    CONST robtarget Target_Nom_Rint_40:=[[-62.519469,-32.68026,0],[0.707106781,0,0,0.707106781],[0,0,0,0],[9E+09,9E+09,9E+09,9E+09,9E+09,9E+09]];
    CONST robtarget Target_Nom_Rint_50:=[[-62.519469,-22.091371,0],[0.707106781,0,0,0.707106781],[0,0,0,0],[9E+09,9E+09,9E+09,9E+09,9E+09,9E+09]];
    CONST robtarget Target_Nom_Rint_60:=[[-87.445335,-22.18424,0],[0.707106781,0,0,0.707106781],[0,0,0,0],[9E+09,9E+09,9E+09,9E+09,9E+09,9E+09]];
    CONST robtarget Target_Nom_Rint_70:=[[-87.50619,-27.43225,0],[0.707106781,0,0,0.707106781],[0,0,0,0],[9E+09,9E+09,9E+09,9E+09,9E+09,9E+09]];
    CONST robtarget Target_Nom_Rint_80:=[[-87.50619,-27.43225,-20],[0.707106781,0,0,0.707106781],[0,0,0,0],[9E+09,9E+09,9E+09,9E+09,9E+09,9E+09]];
    !***********************************************************

    !Dise?o de la parte frontal
    !***********************************************************
    !Punto para acomodar orientaci?n del defector
    CONST robtarget Target_Frente_10:=[[212.749496796,-44.184,-87.888947338],[0.627211375,-0.326505577,-0.326505577,0.627211375],[0,0,0,0],[9E+09,9E+09,9E+09,9E+09,9E+09,9E+09]];
    CONST robtarget Target_Frente_20:=[[196.247119583,-40.184,-39.636157587],[0.428395846,-0.281546356,-0.169146611,0.841782675],[0,0,0,0],[9E+09,9E+09,9E+09,9E+09,9E+09,9E+09]];
    !***********************************************************
    !Dibujo de chip
    CONST robtarget Target_DibChip_10:=[[143.048,-41.184,47.089],[0.595801453,-0.480725183,-0.403998863,0.500708343],[0,0,0,0],[9E+09,9E+09,9E+09,9E+09,9E+09,9E+09]];
    CONST robtarget Target_DibChip_20:=[[123.048,-31.184,47.089],[0.595801453,-0.480725183,-0.403998863,0.500708343],[0,0,0,0],[9E+09,9E+09,9E+09,9E+09,9E+09,9E+09]];
    CONST robtarget Target_DibChip_30:=[[122.19,-34.343,47.089],[0.595801453,-0.480725183,-0.403998863,0.500708343],[0,0,0,0],[9E+09,9E+09,9E+09,9E+09,9E+09,9E+09]];
    CONST robtarget Target_DibChip_40:=[[122.19,-34.343,43.815],[0.595801453,-0.480725183,-0.403998863,0.500708343],[0,0,0,0],[9E+09,9E+09,9E+09,9E+09,9E+09,9E+09]];
    CONST robtarget Target_DibChip_50:=[[122.19,-34.343,47.089],[0.595801453,-0.480725183,-0.403998863,0.500708343],[0,0,0,0],[9E+09,9E+09,9E+09,9E+09,9E+09,9E+09]];
    CONST robtarget Target_DibChip_60:=[[119.685,-42.135,47.089],[0.595801453,-0.480725183,-0.403998863,0.500708343],[0,0,0,0],[9E+09,9E+09,9E+09,9E+09,9E+09,9E+09]];
    CONST robtarget Target_DibChip_70:=[[119.685,-42.135,43.815],[0.595801453,-0.480725183,-0.403998863,0.500708343],[0,0,0,0],[9E+09,9E+09,9E+09,9E+09,9E+09,9E+09]];
    CONST robtarget Target_DibChip_80:=[[119.685,-42.135,47.089],[0.595801453,-0.480725183,-0.403998863,0.500708343],[0,0,0,0],[9E+09,9E+09,9E+09,9E+09,9E+09,9E+09]];
    CONST robtarget Target_DibChip_90:=[[116.675,-49.746,47.089],[0.595801453,-0.480725183,-0.403998863,0.500708343],[0,0,0,0],[9E+09,9E+09,9E+09,9E+09,9E+09,9E+09]];
    CONST robtarget Target_DibChip_100:=[[116.675,-49.746,43.815],[0.595801453,-0.480725183,-0.403998863,0.500708343],[0,0,0,0],[9E+09,9E+09,9E+09,9E+09,9E+09,9E+09]];
    CONST robtarget Target_DibChip_110:=[[116.675,-49.746,47.089],[0.595801453,-0.480725183,-0.403998863,0.500708343],[0,0,0,0],[9E+09,9E+09,9E+09,9E+09,9E+09,9E+09]];
    CONST robtarget Target_DibChip_120:=[[115.333,-52.732,47.089],[0.595801453,-0.480725183,-0.403998863,0.500708343],[0,0,0,0],[9E+09,9E+09,9E+09,9E+09,9E+09,9E+09]];
    CONST robtarget Target_DibChip_130:=[[113.824,-55.86,48.528],[0.595801453,-0.480725183,-0.403998863,0.500708343],[0,0,0,0],[9E+09,9E+09,9E+09,9E+09,9E+09,9E+09]];
    CONST robtarget Target_DibChip_140:=[[113.174,-57.143,52.001],[0.595801453,-0.480725183,-0.403998863,0.500708343],[0,0,0,0],[9E+09,9E+09,9E+09,9E+09,9E+09,9E+09]];
    CONST robtarget Target_DibChip_150:=[[113.174,-57.143,55.275],[0.595801453,-0.480725183,-0.403998863,0.500708343],[0,0,0,0],[9E+09,9E+09,9E+09,9E+09,9E+09,9E+09]];
    CONST robtarget Target_DibChip_160:=[[111.639,-60.035,55.275],[0.595801453,-0.480725183,-0.403998863,0.500708343],[0,0,0,0],[9E+09,9E+09,9E+09,9E+09,9E+09,9E+09]];
    CONST robtarget Target_DibChip_170:=[[113.174,-57.143,55.275],[0.595801453,-0.480725183,-0.403998863,0.500708343],[0,0,0,0],[9E+09,9E+09,9E+09,9E+09,9E+09,9E+09]];
    CONST robtarget Target_DibChip_180:=[[113.174,-57.143,63.46],[0.595801453,-0.480725183,-0.403998863,0.500708343],[0,0,0,0],[9E+09,9E+09,9E+09,9E+09,9E+09,9E+09]];
    CONST robtarget Target_DibChip_190:=[[111.639,-60.035,63.46],[0.595801453,-0.480725183,-0.403998863,0.500708343],[0,0,0,0],[9E+09,9E+09,9E+09,9E+09,9E+09,9E+09]];
    CONST robtarget Target_DibChip_200:=[[113.174,-57.143,63.46],[0.595801453,-0.480725183,-0.403998863,0.500708343],[0,0,0,0],[9E+09,9E+09,9E+09,9E+09,9E+09,9E+09]];
    CONST robtarget Target_DibChip_210:=[[113.174,-57.143,71.646],[0.595801453,-0.480725183,-0.403998863,0.500708343],[0,0,0,0],[9E+09,9E+09,9E+09,9E+09,9E+09,9E+09]];
    CONST robtarget Target_DibChip_220:=[[111.639,-60.035,71.646],[0.595801453,-0.480725183,-0.403998863,0.500708343],[0,0,0,0],[9E+09,9E+09,9E+09,9E+09,9E+09,9E+09]];
    CONST robtarget Target_DibChip_230:=[[113.174,-57.143,71.646],[0.595801453,-0.480725183,-0.403998863,0.500708343],[0,0,0,0],[9E+09,9E+09,9E+09,9E+09,9E+09,9E+09]];
    CONST robtarget Target_DibChip_240:=[[113.174,-57.143,74.92],[0.595801453,-0.480725183,-0.403998863,0.500708343],[0,0,0,0],[9E+09,9E+09,9E+09,9E+09,9E+09,9E+09]];
    CONST robtarget Target_DibChip_250:=[[113.824,-55.86,78.393],[0.595801453,-0.480725183,-0.403998863,0.500708343],[0,0,0,0],[9E+09,9E+09,9E+09,9E+09,9E+09,9E+09]];
    CONST robtarget Target_DibChip_260:=[[115.333,-52.732,79.832],[0.595801453,-0.480725183,-0.403998863,0.500708343],[0,0,0,0],[9E+09,9E+09,9E+09,9E+09,9E+09,9E+09]];
    CONST robtarget Target_DibChip_270:=[[116.675,-49.746,79.832],[0.595801453,-0.480725183,-0.403998863,0.500708343],[0,0,0,0],[9E+09,9E+09,9E+09,9E+09,9E+09,9E+09]];
    CONST robtarget Target_DibChip_280:=[[116.675,-49.746,83.106],[0.595801453,-0.480725183,-0.403998863,0.500708343],[0,0,0,0],[9E+09,9E+09,9E+09,9E+09,9E+09,9E+09]];
    CONST robtarget Target_DibChip_290:=[[116.675,-49.746,79.832],[0.595801453,-0.480725183,-0.403998863,0.500708343],[0,0,0,0],[9E+09,9E+09,9E+09,9E+09,9E+09,9E+09]];
    CONST robtarget Target_DibChip_300:=[[119.685,-42.135,79.832],[0.595801453,-0.480725183,-0.403998863,0.500708343],[0,0,0,0],[9E+09,9E+09,9E+09,9E+09,9E+09,9E+09]];
    CONST robtarget Target_DibChip_310:=[[119.685,-42.135,83.106],[0.595801453,-0.480725183,-0.403998863,0.500708343],[0,0,0,0],[9E+09,9E+09,9E+09,9E+09,9E+09,9E+09]];
    CONST robtarget Target_DibChip_320:=[[119.685,-42.135,79.832],[0.595801453,-0.480725183,-0.403998863,0.500708343],[0,0,0,0],[9E+09,9E+09,9E+09,9E+09,9E+09,9E+09]];
    CONST robtarget Target_DibChip_330:=[[122.19,-34.343,79.832],[0.595801453,-0.480725183,-0.403998863,0.500708343],[0,0,0,0],[9E+09,9E+09,9E+09,9E+09,9E+09,9E+09]];
    CONST robtarget Target_DibChip_340:=[[122.19,-34.343,83.106],[0.595801453,-0.480725183,-0.403998863,0.500708343],[0,0,0,0],[9E+09,9E+09,9E+09,9E+09,9E+09,9E+09]];
    CONST robtarget Target_DibChip_350:=[[122.19,-34.343,79.832],[0.595801453,-0.480725183,-0.403998863,0.500708343],[0,0,0,0],[9E+09,9E+09,9E+09,9E+09,9E+09,9E+09]];
    CONST robtarget Target_DibChip_360:=[[123.048,-31.184,79.832],[0.595801453,-0.480725183,-0.403998863,0.500708343],[0,0,0,0],[9E+09,9E+09,9E+09,9E+09,9E+09,9E+09]];
    CONST robtarget Target_DibChip_370:=[[123.867,-27.809,78.393],[0.595801453,-0.480725183,-0.403998863,0.500708343],[0,0,0,0],[9E+09,9E+09,9E+09,9E+09,9E+09,9E+09]];
    CONST robtarget Target_DibChip_380:=[[124.179,-26.405,74.92],[0.595801453,-0.480725183,-0.403998863,0.500708343],[0,0,0,0],[9E+09,9E+09,9E+09,9E+09,9E+09,9E+09]];
    CONST robtarget Target_DibChip_390:=[[124.179,-26.405,71.646],[0.595801453,-0.480725183,-0.403998863,0.500708343],[0,0,0,0],[9E+09,9E+09,9E+09,9E+09,9E+09,9E+09]];
    CONST robtarget Target_DibChip_400:=[[124.829,-23.196,71.646],[0.595801453,-0.480725183,-0.403998863,0.500708343],[0,0,0,0],[9E+09,9E+09,9E+09,9E+09,9E+09,9E+09]];
    CONST robtarget Target_DibChip_410:=[[124.179,-26.405,71.646],[0.595801453,-0.480725183,-0.403998863,0.500708343],[0,0,0,0],[9E+09,9E+09,9E+09,9E+09,9E+09,9E+09]];
    CONST robtarget Target_DibChip_420:=[[124.179,-26.405,63.46],[0.595801453,-0.480725183,-0.403998863,0.500708343],[0,0,0,0],[9E+09,9E+09,9E+09,9E+09,9E+09,9E+09]];
    CONST robtarget Target_DibChip_430:=[[124.829,-23.196,63.46],[0.595801453,-0.480725183,-0.403998863,0.500708343],[0,0,0,0],[9E+09,9E+09,9E+09,9E+09,9E+09,9E+09]];
    CONST robtarget Target_DibChip_440:=[[124.179,-26.405,63.46],[0.595801453,-0.480725183,-0.403998863,0.500708343],[0,0,0,0],[9E+09,9E+09,9E+09,9E+09,9E+09,9E+09]];
    CONST robtarget Target_DibChip_450:=[[124.179,-26.405,55.275],[0.595801453,-0.480725183,-0.403998863,0.500708343],[0,0,0,0],[9E+09,9E+09,9E+09,9E+09,9E+09,9E+09]];
    CONST robtarget Target_DibChip_460:=[[124.829,-23.196,55.275],[0.595801453,-0.480725183,-0.403998863,0.500708343],[0,0,0,0],[9E+09,9E+09,9E+09,9E+09,9E+09,9E+09]];
    CONST robtarget Target_DibChip_470:=[[124.179,-26.405,55.275],[0.595801453,-0.480725183,-0.403998863,0.500708343],[0,0,0,0],[9E+09,9E+09,9E+09,9E+09,9E+09,9E+09]];
    CONST robtarget Target_DibChip_480:=[[124.179,-26.405,52.001],[0.595801453,-0.480725183,-0.403998863,0.500708343],[0,0,0,0],[9E+09,9E+09,9E+09,9E+09,9E+09,9E+09]];
    CONST robtarget Target_DibChip_490:=[[123.867,-27.809,48.528],[0.595801453,-0.480725183,-0.403998863,0.500708343],[0,0,0,0],[9E+09,9E+09,9E+09,9E+09,9E+09,9E+09]];
    CONST robtarget Target_DibChip_500:=[[123.048,-31.184,47.089],[0.595801453,-0.480725183,-0.403998863,0.500708343],[0,0,0,0],[9E+09,9E+09,9E+09,9E+09,9E+09,9E+09]];
    CONST robtarget Target_DibChip_510:=[[143.048,-41.184,47.089],[0.595801453,-0.480725183,-0.403998863,0.500708343],[0,0,0,0],[9E+09,9E+09,9E+09,9E+09,9E+09,9E+09]];
    CONST robtarget Target_DibChip_520:=[[142.629,-42.767,53.638],[0.595801453,-0.480725183,-0.403998863,0.500708343],[-1,0,-1,0],[9E+09,9E+09,9E+09,9E+09,9E+09,9E+09]];
    CONST robtarget Target_DibChip_530:=[[122.629,-32.767,53.638],[0.595801453,-0.480725183,-0.403998863,0.500708343],[-1,0,-1,0],[9E+09,9E+09,9E+09,9E+09,9E+09,9E+09]];
    CONST robtarget Target_DibChip_540:=[[116.014,-51.243,53.638],[0.595801453,-0.480725183,-0.403998863,0.500708343],[-1,0,-1,0],[9E+09,9E+09,9E+09,9E+09,9E+09,9E+09]];
    CONST robtarget Target_DibChip_550:=[[116.014,-51.243,73.283],[0.595801453,-0.480725183,-0.403998863,0.500708343],[-1,0,-1,0],[9E+09,9E+09,9E+09,9E+09,9E+09,9E+09]];
    CONST robtarget Target_DibChip_560:=[[122.629,-32.767,73.283],[0.595801453,-0.480725183,-0.403998863,0.500708343],[-1,0,-1,0],[9E+09,9E+09,9E+09,9E+09,9E+09,9E+09]];
    CONST robtarget Target_DibChip_570:=[[122.629,-32.767,53.638],[0.595801453,-0.480725183,-0.403998863,0.500708343],[-1,0,-1,0],[9E+09,9E+09,9E+09,9E+09,9E+09,9E+09]];
    CONST robtarget Target_DibChip_580:=[[142.629,-42.767,53.638],[0.595801453,-0.480725183,-0.403998863,0.500708343],[0,0,0,0],[9E+09,9E+09,9E+09,9E+09,9E+09,9E+09]];
    !***********************************************************
    !Dibujo primer cuadrante de letrero frontal
    CONST robtarget Target_LetFron1_10:=[[106.389,-99.587,43.347],[0.680036541,-0.521810391,-0.313535314,0.408607177],[0,0,0,0],[9E+09,9E+09,9E+09,9E+09,9E+09,9E+09]];
    CONST robtarget Target_LetFron1_20:=[[96.389,-79.587,43.347],[0.680036541,-0.521810391,-0.313535314,0.408607177],[0,0,0,0],[9E+09,9E+09,9E+09,9E+09,9E+09,9E+09]];
    CONST robtarget Target_LetFron1_30:=[[96.389,-79.587,57.11],[0.680036541,-0.521810391,-0.313535314,0.408607177],[0,0,0,0],[9E+09,9E+09,9E+09,9E+09,9E+09,9E+09]];
    CONST robtarget Target_LetFron1_40:=[[91.42,-85.249,57.11],[0.680036541,-0.521810391,-0.313535314,0.408607177],[0,0,0,0],[9E+09,9E+09,9E+09,9E+09,9E+09,9E+09]];
    CONST robtarget Target_LetFron1_50:=[[101.42,-105.249,57.11],[0.680036541,-0.521810391,-0.313535314,0.408607177],[0,0,0,0],[9E+09,9E+09,9E+09,9E+09,9E+09,9E+09]];
    CONST robtarget Target_LetFron1_60:=[[100.543,-106.18,48.283],[0.680036541,-0.521810391,-0.313535314,0.408607177],[0,0,0,0],[9E+09,9E+09,9E+09,9E+09,9E+09,9E+09]];
    CONST robtarget Target_LetFron1_70:=[[90.543,-86.18,48.283],[0.680036541,-0.521810391,-0.313535314,0.408607177],[0,0,0,0],[9E+09,9E+09,9E+09,9E+09,9E+09,9E+09]];
    CONST robtarget Target_LetFron1_80:=[[86.36,-90.371,47.26],[0.680036541,-0.521810391,-0.313535314,0.408607177],[0,0,0,0],[9E+09,9E+09,9E+09,9E+09,9E+09,9E+09]];
    CONST robtarget Target_LetFron1_90:=[[85.516,-91.17,49.426],[0.680036541,-0.521810391,-0.313535314,0.408607177],[0,0,0,0],[9E+09,9E+09,9E+09,9E+09,9E+09,9E+09]];
    CONST robtarget Target_LetFron1_100:=[[85.516,-91.17,53.546],[0.680036541,-0.521810391,-0.313535314,0.408607177],[0,0,0,0],[9E+09,9E+09,9E+09,9E+09,9E+09,9E+09]];
    CONST robtarget Target_LetFron1_110:=[[85.516,-91.17,57.11],[0.680036541,-0.521810391,-0.313535314,0.408607177],[0,0,0,0],[9E+09,9E+09,9E+09,9E+09,9E+09,9E+09]];
    CONST robtarget Target_LetFron1_120:=[[86.479,-90.257,57.403],[0.680036541,-0.521810391,-0.313535314,0.408607177],[0,0,0,0],[9E+09,9E+09,9E+09,9E+09,9E+09,9E+09]];
    CONST robtarget Target_LetFron1_130:=[[86.771,-89.977,56.211],[0.680036541,-0.521810391,-0.313535314,0.408607177],[0,0,0,0],[9E+09,9E+09,9E+09,9E+09,9E+09,9E+09]];
    CONST robtarget Target_LetFron1_140:=[[88.867,-87.907,57.403],[0.680036541,-0.521810391,-0.313535314,0.408607177],[0,0,0,0],[9E+09,9E+09,9E+09,9E+09,9E+09,9E+09]];
    CONST robtarget Target_LetFron1_150:=[[90.326,-86.408,56.683],[0.680036541,-0.521810391,-0.313535314,0.408607177],[0,0,0,0],[9E+09,9E+09,9E+09,9E+09,9E+09,9E+09]];
    CONST robtarget Target_LetFron1_160:=[[90.899,-85.804,54.727],[0.680036541,-0.521810391,-0.313535314,0.408607177],[0,0,0,0],[9E+09,9E+09,9E+09,9E+09,9E+09,9E+09]];
    CONST robtarget Target_LetFron1_170:=[[89.983,-86.764,52.388],[0.680036541,-0.521810391,-0.313535314,0.408607177],[0,0,0,0],[9E+09,9E+09,9E+09,9E+09,9E+09,9E+09]];
    CONST robtarget Target_LetFron1_180:=[[88.854,-87.92,51.608],[0.680036541,-0.521810391,-0.313535314,0.408607177],[0,0,0,0],[9E+09,9E+09,9E+09,9E+09,9E+09,9E+09]];
    CONST robtarget Target_LetFron1_190:=[[86.884,-89.867,51.398],[0.680036541,-0.521810391,-0.313535314,0.408607177],[0,0,0,0],[9E+09,9E+09,9E+09,9E+09,9E+09,9E+09]];
    CONST robtarget Target_LetFron1_200:=[[106.884,-109.867,51.398],[0.680036541,-0.521810391,-0.313535314,0.408607177],[0,0,0,0],[9E+09,9E+09,9E+09,9E+09,9E+09,9E+09]];
    CONST robtarget Target_LetFron1_210:=[[103.236,-113.256,41.93],[0.680036541,-0.521810391,-0.313535314,0.408607177],[0,0,0,0],[9E+09,9E+09,9E+09,9E+09,9E+09,9E+09]];
    CONST robtarget Target_LetFron1_220:=[[83.236,-93.256,41.93],[0.680036541,-0.521810391,-0.313535314,0.408607177],[0,0,0,0],[9E+09,9E+09,9E+09,9E+09,9E+09,9E+09]];
    CONST robtarget Target_LetFron1_230:=[[83.236,-93.256,57.358],[0.680036541,-0.521810391,-0.313535314,0.408607177],[0,0,0,0],[9E+09,9E+09,9E+09,9E+09,9E+09,9E+09]];
    CONST robtarget Target_LetFron1_240:=[[82.597,-93.823,57.628],[0.680036541,-0.521810391,-0.313535314,0.408607177],[0,0,0,0],[9E+09,9E+09,9E+09,9E+09,9E+09,9E+09]];
    CONST robtarget Target_LetFron1_250:=[[82.208,-94.164,56.818],[0.680036541,-0.521810391,-0.313535314,0.408607177],[0,0,0,0],[9E+09,9E+09,9E+09,9E+09,9E+09,9E+09]];
    CONST robtarget Target_LetFron1_260:=[[80.629,-95.519,57.358],[0.680036541,-0.521810391,-0.313535314,0.408607177],[0,0,0,0],[9E+09,9E+09,9E+09,9E+09,9E+09,9E+09]];
    CONST robtarget Target_LetFron1_270:=[[78.563,-97.226,56.975],[0.680036541,-0.521810391,-0.313535314,0.408607177],[0,0,0,0],[9E+09,9E+09,9E+09,9E+09,9E+09,9E+09]];
    CONST robtarget Target_LetFron1_280:=[[77.179,-98.328,55.611],[0.680036541,-0.521810391,-0.313535314,0.408607177],[0,0,0,0],[9E+09,9E+09,9E+09,9E+09,9E+09,9E+09]];
    CONST robtarget Target_LetFron1_290:=[[76.653,-98.738,54.322],[0.680036541,-0.521810391,-0.313535314,0.408607177],[0,0,0,0],[9E+09,9E+09,9E+09,9E+09,9E+09,9E+09]];
    CONST robtarget Target_LetFron1_300:=[[76.4,-98.935,53.152],[0.680036541,-0.521810391,-0.313535314,0.408607177],[0,0,0,0],[9E+09,9E+09,9E+09,9E+09,9E+09,9E+09]];
    CONST robtarget Target_LetFron1_310:=[[76.315,-99,51.196],[0.680036541,-0.521810391,-0.313535314,0.408607177],[0,0,0,0],[9E+09,9E+09,9E+09,9E+09,9E+09,9E+09]];
    CONST robtarget Target_LetFron1_320:=[[76.475,-98.876,49.614],[0.680036541,-0.521810391,-0.313535314,0.408607177],[0,0,0,0],[9E+09,9E+09,9E+09,9E+09,9E+09,9E+09]];
    CONST robtarget Target_LetFron1_330:=[[77.102,-98.388,48.13],[0.680036541,-0.521810391,-0.313535314,0.408607177],[0,0,0,0],[9E+09,9E+09,9E+09,9E+09,9E+09,9E+09]];
    CONST robtarget Target_LetFron1_340:=[[78.458,-97.311,46.893],[0.680036541,-0.521810391,-0.313535314,0.408607177],[0,0,0,0],[9E+09,9E+09,9E+09,9E+09,9E+09,9E+09]];
    CONST robtarget Target_LetFron1_350:=[[79.625,-96.358,46.72],[0.680036541,-0.521810391,-0.313535314,0.408607177],[0,0,0,0],[9E+09,9E+09,9E+09,9E+09,9E+09,9E+09]];
    CONST robtarget Target_LetFron1_360:=[[80.34,-95.763,46.9],[0.680036541,-0.521810391,-0.313535314,0.408607177],[0,0,0,0],[9E+09,9E+09,9E+09,9E+09,9E+09,9E+09]];
    CONST robtarget Target_LetFron1_370:=[[81.139,-95.086,47.294],[0.680036541,-0.521810391,-0.313535314,0.408607177],[0,0,0,0],[9E+09,9E+09,9E+09,9E+09,9E+09,9E+09]];
    CONST robtarget Target_LetFron1_380:=[[81.783,-94.533,47.71],[0.680036541,-0.521810391,-0.313535314,0.408607177],[0,0,0,0],[9E+09,9E+09,9E+09,9E+09,9E+09,9E+09]];
    CONST robtarget Target_LetFron1_390:=[[101.783,-114.533,47.71],[0.680036541,-0.521810391,-0.313535314,0.408607177],[0,0,0,0],[9E+09,9E+09,9E+09,9E+09,9E+09,9E+09]];
    CONST robtarget Target_LetFron1_400:=[[84.525,-120.354,49.262],[0.680036541,-0.521810391,-0.313535314,0.408607177],[0,0,0,0],[9E+09,9E+09,9E+09,9E+09,9E+09,9E+09]];
    CONST robtarget Target_LetFron1_410:=[[74.525,-100.354,49.262],[0.680036541,-0.521810391,-0.313535314,0.408607177],[0,0,0,0],[9E+09,9E+09,9E+09,9E+09,9E+09,9E+09]];
    CONST robtarget Target_LetFron1_420:=[[74.946,-100.041,50.585],[0.680036541,-0.521810391,-0.313535314,0.408607177],[0,0,0,0],[9E+09,9E+09,9E+09,9E+09,9E+09,9E+09]];
    CONST robtarget Target_LetFron1_430:=[[75.03,-99.978,51.668],[0.680036541,-0.521810391,-0.313535314,0.408607177],[0,0,0,0],[9E+09,9E+09,9E+09,9E+09,9E+09,9E+09]];
    CONST robtarget Target_LetFron1_440:=[[75.03,-99.978,53.347],[0.680036541,-0.521810391,-0.313535314,0.408607177],[0,0,0,0],[9E+09,9E+09,9E+09,9E+09,9E+09,9E+09]];
    CONST robtarget Target_LetFron1_450:=[[74.718,-100.211,54.659],[0.680036541,-0.521810391,-0.313535314,0.408607177],[0,0,0,0],[9E+09,9E+09,9E+09,9E+09,9E+09,9E+09]];
    CONST robtarget Target_LetFron1_460:=[[73.992,-100.748,56.053],[0.680036541,-0.521810391,-0.313535314,0.408607177],[0,0,0,0],[9E+09,9E+09,9E+09,9E+09,9E+09,9E+09]];
    CONST robtarget Target_LetFron1_470:=[[72.976,-101.487,56.998],[0.680036541,-0.521810391,-0.313535314,0.408607177],[0,0,0,0],[9E+09,9E+09,9E+09,9E+09,9E+09,9E+09]];
    CONST robtarget Target_LetFron1_480:=[[71.366,-102.625,57.403],[0.680036541,-0.521810391,-0.313535314,0.408607177],[0,0,0,0],[9E+09,9E+09,9E+09,9E+09,9E+09,9E+09]];
    CONST robtarget Target_LetFron1_490:=[[69.446,-103.934,56.968],[0.680036541,-0.521810391,-0.313535314,0.408607177],[0,0,0,0],[9E+09,9E+09,9E+09,9E+09,9E+09,9E+09]];
    CONST robtarget Target_LetFron1_500:=[[68.289,-104.698,55.935],[0.680036541,-0.521810391,-0.313535314,0.408607177],[0,0,0,0],[9E+09,9E+09,9E+09,9E+09,9E+09,9E+09]];
    CONST robtarget Target_LetFron1_510:=[[67.489,-105.215,54.419],[0.680036541,-0.521810391,-0.313535314,0.408607177],[0,0,0,0],[9E+09,9E+09,9E+09,9E+09,9E+09,9E+09]];
    CONST robtarget Target_LetFron1_520:=[[67.135,-105.441,53.002],[0.680036541,-0.521810391,-0.313535314,0.408607177],[0,0,0,0],[9E+09,9E+09,9E+09,9E+09,9E+09,9E+09]];
    CONST robtarget Target_LetFron1_530:=[[67.135,-105.441,50.753],[0.680036541,-0.521810391,-0.313535314,0.408607177],[0,0,0,0],[9E+09,9E+09,9E+09,9E+09,9E+09,9E+09]];
    CONST robtarget Target_LetFron1_540:=[[67.609,-105.138,49.082],[0.680036541,-0.521810391,-0.313535314,0.408607177],[0,0,0,0],[9E+09,9E+09,9E+09,9E+09,9E+09,9E+09]];
    CONST robtarget Target_LetFron1_550:=[[67.924,-104.935,48.317],[0.680036541,-0.521810391,-0.313535314,0.408607177],[0,0,0,0],[9E+09,9E+09,9E+09,9E+09,9E+09,9E+09]];
    CONST robtarget Target_LetFron1_560:=[[68.928,-104.278,47.327],[0.680036541,-0.521810391,-0.313535314,0.408607177],[0,0,0,0],[9E+09,9E+09,9E+09,9E+09,9E+09,9E+09]];
    CONST robtarget Target_LetFron1_570:=[[69.801,-103.696,46.821],[0.680036541,-0.521810391,-0.313535314,0.408607177],[0,0,0,0],[9E+09,9E+09,9E+09,9E+09,9E+09,9E+09]];
    CONST robtarget Target_LetFron1_580:=[[70.496,-103.225,46.72],[0.680036541,-0.521810391,-0.313535314,0.408607177],[0,0,0,0],[9E+09,9E+09,9E+09,9E+09,9E+09,9E+09]];
    CONST robtarget Target_LetFron1_590:=[[71.729,-102.372,46.72],[0.680036541,-0.521810391,-0.313535314,0.408607177],[0,0,0,0],[9E+09,9E+09,9E+09,9E+09,9E+09,9E+09]];
    CONST robtarget Target_LetFron1_600:=[[72.47,-101.849,46.938],[0.680036541,-0.521810391,-0.313535314,0.408607177],[0,0,0,0],[9E+09,9E+09,9E+09,9E+09,9E+09,9E+09]];
    CONST robtarget Target_LetFron1_610:=[[73.401,-101.179,47.59],[0.680036541,-0.521810391,-0.313535314,0.408607177],[0,0,0,0],[9E+09,9E+09,9E+09,9E+09,9E+09,9E+09]];
    CONST robtarget Target_LetFron1_620:=[[74.188,-100.604,48.437],[0.680036541,-0.521810391,-0.313535314,0.408607177],[0,0,0,0],[9E+09,9E+09,9E+09,9E+09,9E+09,9E+09]];
    CONST robtarget Target_LetFron1_630:=[[74.525,-100.354,49.262],[0.680036541,-0.521810391,-0.313535314,0.408607177],[0,0,0,0],[9E+09,9E+09,9E+09,9E+09,9E+09,9E+09]];
    CONST robtarget Target_LetFron1_640:=[[84.188,-120.604,48.437],[0.680036541,-0.521810391,-0.313535314,0.408607177],[0,0,0,0],[9E+09,9E+09,9E+09,9E+09,9E+09,9E+09]];
    CONST robtarget Target_LetFron1_650:=[[74.265,-127.215,57.11],[0.680036541,-0.521810391,-0.313535314,0.408607177],[0,0,0,0],[9E+09,9E+09,9E+09,9E+09,9E+09,9E+09]];
    CONST robtarget Target_LetFron1_660:=[[64.265,-107.215,57.11],[0.680036541,-0.521810391,-0.313535314,0.408607177],[0,0,0,0],[9E+09,9E+09,9E+09,9E+09,9E+09,9E+09]];
    CONST robtarget Target_LetFron1_670:=[[64.496,-107.076,46.866],[0.680036541,-0.521810391,-0.313535314,0.408607177],[0,0,0,0],[9E+09,9E+09,9E+09,9E+09,9E+09,9E+09]];
    CONST robtarget Target_LetFron1_680:=[[63.362,-107.751,47.897],[0.680036541,-0.521810391,-0.313535314,0.408607177],[0,0,0,0],[9E+09,9E+09,9E+09,9E+09,9E+09,9E+09]];
    CONST robtarget Target_LetFron1_690:=[[61.942,-108.574,46.863],[0.680036541,-0.521810391,-0.313535314,0.408607177],[0,0,0,0],[9E+09,9E+09,9E+09,9E+09,9E+09,9E+09]];
    CONST robtarget Target_LetFron1_700:=[[60.609,-109.323,46.758],[0.680036541,-0.521810391,-0.313535314,0.408607177],[0,0,0,0],[9E+09,9E+09,9E+09,9E+09,9E+09,9E+09]];
    CONST robtarget Target_LetFron1_710:=[[70.609,-129.323,46.758],[0.680036541,-0.521810391,-0.313535314,0.408607177],[0,0,0,0],[9E+09,9E+09,9E+09,9E+09,9E+09,9E+09]];
    CONST robtarget Target_LetFron1_720:=[[69.365,-120.003,48.283],[0.680036541,-0.521810391,-0.313535314,0.408607177],[0,0,0,0],[9E+09,9E+09,9E+09,9E+09,9E+09,9E+09]];
    CONST robtarget Target_LetFron1_730:=[[59.365,-110.003,48.283],[0.680036541,-0.521810391,-0.313535314,0.408607177],[0,0,0,0],[9E+09,9E+09,9E+09,9E+09,9E+09,9E+09]];
    CONST robtarget Target_LetFron1_740:=[[54.346,-112.568,46.99],[0.680036541,-0.521810391,-0.313535314,0.408607177],[0,0,0,0],[9E+09,9E+09,9E+09,9E+09,9E+09,9E+09]];
    CONST robtarget Target_LetFron1_750:=[[53.304,-113.065,48.055],[0.680036541,-0.521810391,-0.313535314,0.408607177],[0,0,0,0],[9E+09,9E+09,9E+09,9E+09,9E+09,9E+09]];
    CONST robtarget Target_LetFron1_760:=[[53.039,-113.189,48.872],[0.680036541,-0.521810391,-0.313535314,0.408607177],[0,0,0,0],[9E+09,9E+09,9E+09,9E+09,9E+09,9E+09]];
    CONST robtarget Target_LetFron1_770:=[[53.039,-113.189,49.981],[0.680036541,-0.521810391,-0.313535314,0.408607177],[0,0,0,0],[9E+09,9E+09,9E+09,9E+09,9E+09,9E+09]];
    CONST robtarget Target_LetFron1_780:=[[53.039,-113.189,57.11],[0.680036541,-0.521810391,-0.313535314,0.408607177],[0,0,0,0],[9E+09,9E+09,9E+09,9E+09,9E+09,9E+09]];
    CONST robtarget Target_LetFron1_790:=[[54.238,-112.62,57.403],[0.680036541,-0.521810391,-0.313535314,0.408607177],[0,0,0,0],[9E+09,9E+09,9E+09,9E+09,9E+09,9E+09]];
    CONST robtarget Target_LetFron1_800:=[[54.717,-112.388,56.293],[0.680036541,-0.521810391,-0.313535314,0.408607177],[0,0,0,0],[9E+09,9E+09,9E+09,9E+09,9E+09,9E+09]];
    CONST robtarget Target_LetFron1_810:=[[56.663,-111.42,57.335],[0.680036541,-0.521810391,-0.313535314,0.408607177],[0,0,0,0],[9E+09,9E+09,9E+09,9E+09,9E+09,9E+09]];
    CONST robtarget Target_LetFron1_820:=[[58.249,-110.599,57.223],[0.680036541,-0.521810391,-0.313535314,0.408607177],[0,0,0,0],[9E+09,9E+09,9E+09,9E+09,9E+09,9E+09]];
    CONST robtarget Target_LetFron1_830:=[[59.332,-110.021,56.436],[0.680036541,-0.521810391,-0.313535314,0.408607177],[0,0,0,0],[9E+09,9E+09,9E+09,9E+09,9E+09,9E+09]];
    CONST robtarget Target_LetFron1_840:=[[59.82,-109.757,55.131],[0.680036541,-0.521810391,-0.313535314,0.408607177],[0,0,0,0],[9E+09,9E+09,9E+09,9E+09,9E+09,9E+09]];
    CONST robtarget Target_LetFron1_850:=[[59.82,-109.757,54.254],[0.680036541,-0.521810391,-0.313535314,0.408607177],[0,0,0,0],[9E+09,9E+09,9E+09,9E+09,9E+09,9E+09]];
    CONST robtarget Target_LetFron1_860:=[[59.431,-109.968,53.002],[0.680036541,-0.521810391,-0.313535314,0.408607177],[0,0,0,0],[9E+09,9E+09,9E+09,9E+09,9E+09,9E+09]];
    CONST robtarget Target_LetFron1_870:=[[58.261,-110.592,52.08],[0.680036541,-0.521810391,-0.313535314,0.408607177],[0,0,0,0],[9E+09,9E+09,9E+09,9E+09,9E+09,9E+09]];
    CONST robtarget Target_LetFron1_880:=[[56.569,-111.467,51.443],[0.680036541,-0.521810391,-0.313535314,0.408607177],[0,0,0,0],[9E+09,9E+09,9E+09,9E+09,9E+09,9E+09]];
    CONST robtarget Target_LetFron1_890:=[[54.744,-112.375,51.398],[0.680036541,-0.521810391,-0.313535314,0.408607177],[0,0,0,0],[9E+09,9E+09,9E+09,9E+09,9E+09,9E+09]];
    CONST robtarget Target_LetFron1_900:=[[64.744,-122.375,51.398],[0.680036541,-0.521810391,-0.313535314,0.408607177],[0,0,0,0],[9E+09,9E+09,9E+09,9E+09,9E+09,9E+09]];
    CONST robtarget Target_LetFron1_910:=[[55.006,-126.617,56.155],[0.680036541,-0.521810391,-0.313535314,0.408607177],[0,0,0,0],[9E+09,9E+09,9E+09,9E+09,9E+09,9E+09]];
    CONST robtarget Target_LetFron1_920:=[[45.006,-116.617,56.155],[0.680036541,-0.521810391,-0.313535314,0.408607177],[0,0,0,0],[9E+09,9E+09,9E+09,9E+09,9E+09,9E+09]];
    CONST robtarget Target_LetFron1_930:=[[49.551,-114.759,56.443],[0.680036541,-0.521810391,-0.313535314,0.408607177],[0,0,0,0],[9E+09,9E+09,9E+09,9E+09,9E+09,9E+09]];
    CONST robtarget Target_LetFron1_940:=[[49.967,-114.579,51.567],[0.680036541,-0.521810391,-0.313535314,0.408607177],[0,0,0,0],[9E+09,9E+09,9E+09,9E+09,9E+09,9E+09]];
    CONST robtarget Target_LetFron1_950:=[[49.915,-114.601,46.99],[0.680036541,-0.521810391,-0.313535314,0.408607177],[0,0,0,0],[9E+09,9E+09,9E+09,9E+09,9E+09,9E+09]];
    CONST robtarget Target_LetFron1_960:=[[49.895,-114.61,45.281],[0.680036541,-0.521810391,-0.313535314,0.408607177],[0,0,0,0],[9E+09,9E+09,9E+09,9E+09,9E+09,9E+09]];
    CONST robtarget Target_LetFron1_970:=[[49.915,-114.601,46.99],[0.680036541,-0.521810391,-0.313535314,0.408607177],[0,0,0,0],[9E+09,9E+09,9E+09,9E+09,9E+09,9E+09]];
    CONST robtarget Target_LetFron1_980:=[[51.457,-113.917,47.215],[0.680036541,-0.521810391,-0.313535314,0.408607177],[0,0,0,0],[9E+09,9E+09,9E+09,9E+09,9E+09,9E+09]];
    CONST robtarget Target_LetFron1_990:=[[45.111,-116.576,46.99],[0.680036541,-0.521810391,-0.313535314,0.408607177],[0,0,0,0],[9E+09,9E+09,9E+09,9E+09,9E+09,9E+09]];
    CONST robtarget Target_LetFron1_1000:=[[55.111,-136.576,46.99],[0.680036541,-0.521810391,-0.313535314,0.408607177],[0,0,0,0],[9E+09,9E+09,9E+09,9E+09,9E+09,9E+09]];
    CONST robtarget Target_LetFron1_1010:=[[52.243,-137.646,47.59],[0.680036541,-0.521810391,-0.313535314,0.408607177],[0,0,0,0],[9E+09,9E+09,9E+09,9E+09,9E+09,9E+09]];
    CONST robtarget Target_LetFron1_1020:=[[42.243,-117.646,47.59],[0.680036541,-0.521810391,-0.313535314,0.408607177],[0,0,0,0],[9E+09,9E+09,9E+09,9E+09,9E+09,9E+09]];
    CONST robtarget Target_LetFron1_1030:=[[43.159,-117.313,48.437],[0.680036541,-0.521810391,-0.313535314,0.408607177],[0,0,0,0],[9E+09,9E+09,9E+09,9E+09,9E+09,9E+09]];
    CONST robtarget Target_LetFron1_1040:=[[43.749,-117.094,49.674],[0.680036541,-0.521810391,-0.313535314,0.408607177],[0,0,0,0],[9E+09,9E+09,9E+09,9E+09,9E+09,9E+09]];
    CONST robtarget Target_LetFron1_1050:=[[44.142,-116.946,51.083],[0.680036541,-0.521810391,-0.313535314,0.408607177],[0,0,0,0],[9E+09,9E+09,9E+09,9E+09,9E+09,9E+09]];
    CONST robtarget Target_LetFron1_1060:=[[44.142,-116.946,52.253],[0.680036541,-0.521810391,-0.313535314,0.408607177],[0,0,0,0],[9E+09,9E+09,9E+09,9E+09,9E+09,9E+09]];
    CONST robtarget Target_LetFron1_1070:=[[44.005,-116.998,53.771],[0.680036541,-0.521810391,-0.313535314,0.408607177],[0,0,0,0],[9E+09,9E+09,9E+09,9E+09,9E+09,9E+09]];
    CONST robtarget Target_LetFron1_1080:=[[43.595,-117.152,55.041],[0.680036541,-0.521810391,-0.313535314,0.408607177],[0,0,0,0],[9E+09,9E+09,9E+09,9E+09,9E+09,9E+09]];
    CONST robtarget Target_LetFron1_1090:=[[42.708,-117.478,56.391],[0.680036541,-0.521810391,-0.313535314,0.408607177],[0,0,0,0],[9E+09,9E+09,9E+09,9E+09,9E+09,9E+09]];
    CONST robtarget Target_LetFron1_1100:=[[41.423,-117.937,57.2],[0.680036541,-0.521810391,-0.313535314,0.408607177],[0,0,0,0],[9E+09,9E+09,9E+09,9E+09,9E+09,9E+09]];
    CONST robtarget Target_LetFron1_1110:=[[39.885,-118.466,57.403],[0.680036541,-0.521810391,-0.313535314,0.408607177],[0,0,0,0],[9E+09,9E+09,9E+09,9E+09,9E+09,9E+09]];
    CONST robtarget Target_LetFron1_1120:=[[38.497,-118.924,57.24],[0.680036541,-0.521810391,-0.313535314,0.408607177],[0,0,0,0],[9E+09,9E+09,9E+09,9E+09,9E+09,9E+09]];
    CONST robtarget Target_LetFron1_1130:=[[37.318,-119.299,56.751],[0.680036541,-0.521810391,-0.313535314,0.408607177],[0,0,0,0],[9E+09,9E+09,9E+09,9E+09,9E+09,9E+09]];
    CONST robtarget Target_LetFron1_1140:=[[36.028,-119.695,55.664],[0.680036541,-0.521810391,-0.313535314,0.408607177],[0,0,0,0],[9E+09,9E+09,9E+09,9E+09,9E+09,9E+09]];
    CONST robtarget Target_LetFron1_1150:=[[35.238,-119.93,53.999],[0.680036541,-0.521810391,-0.313535314,0.408607177],[0,0,0,0],[9E+09,9E+09,9E+09,9E+09,9E+09,9E+09]];
    CONST robtarget Target_LetFron1_1160:=[[35.036,-119.989,52.425],[0.680036541,-0.521810391,-0.313535314,0.408607177],[0,0,0,0],[9E+09,9E+09,9E+09,9E+09,9E+09,9E+09]];
    CONST robtarget Target_LetFron1_1170:=[[35.036,-119.989,51.301],[0.680036541,-0.521810391,-0.313535314,0.408607177],[0,0,0,0],[9E+09,9E+09,9E+09,9E+09,9E+09,9E+09]];
    CONST robtarget Target_LetFron1_1180:=[[35.216,-119.937,49.831],[0.680036541,-0.521810391,-0.313535314,0.408607177],[0,0,0,0],[9E+09,9E+09,9E+09,9E+09,9E+09,9E+09]];
    CONST robtarget Target_LetFron1_1190:=[[35.935,-119.723,48.317],[0.680036541,-0.521810391,-0.313535314,0.408607177],[0,0,0,0],[9E+09,9E+09,9E+09,9E+09,9E+09,9E+09]];
    CONST robtarget Target_LetFron1_1200:=[[36.76,-119.473,47.53],[0.680036541,-0.521810391,-0.313535314,0.408607177],[0,0,0,0],[9E+09,9E+09,9E+09,9E+09,9E+09,9E+09]];
    CONST robtarget Target_LetFron1_1210:=[[37.712,-119.176,46.923],[0.680036541,-0.521810391,-0.313535314,0.408607177],[0,0,0,0],[9E+09,9E+09,9E+09,9E+09,9E+09,9E+09]];
    CONST robtarget Target_LetFron1_1220:=[[38.882,-118.799,46.72],[0.680036541,-0.521810391,-0.313535314,0.408607177],[0,0,0,0],[9E+09,9E+09,9E+09,9E+09,9E+09,9E+09]];
    CONST robtarget Target_LetFron1_1230:=[[39.807,-118.492,46.72],[0.680036541,-0.521810391,-0.313535314,0.408607177],[0,0,0,0],[9E+09,9E+09,9E+09,9E+09,9E+09,9E+09]];
    CONST robtarget Target_LetFron1_1240:=[[41.161,-118.029,46.938],[0.680036541,-0.521810391,-0.313535314,0.408607177],[0,0,0,0],[9E+09,9E+09,9E+09,9E+09,9E+09,9E+09]];
    CONST robtarget Target_LetFron1_1250:=[[42.243,-117.646,47.59],[0.680036541,-0.521810391,-0.313535314,0.408607177],[0,0,0,0],[9E+09,9E+09,9E+09,9E+09,9E+09,9E+09]];
    CONST robtarget Target_LetFron1_1260:=[[52.243,-137.646,47.59],[0.680036541,-0.521810391,-0.313535314,0.408607177],[0,0,0,0],[9E+09,9E+09,9E+09,9E+09,9E+09,9E+09]];
    CONST robtarget Target_LetFron1_1270:=[[41.785,-140.891,57.11],[0.680036541,-0.521810391,-0.313535314,0.408607177],[0,0,0,0],[9E+09,9E+09,9E+09,9E+09,9E+09,9E+09]];
    CONST robtarget Target_LetFron1_1280:=[[31.785,-120.891,57.11],[0.680036541,-0.521810391,-0.313535314,0.408607177],[0,0,0,0],[9E+09,9E+09,9E+09,9E+09,9E+09,9E+09]];
    CONST robtarget Target_LetFron1_1290:=[[32.046,-120.822,46.866],[0.680036541,-0.521810391,-0.313535314,0.408607177],[0,0,0,0],[9E+09,9E+09,9E+09,9E+09,9E+09,9E+09]];
    CONST robtarget Target_LetFron1_1300:=[[30.958,-121.106,48.07],[0.680036541,-0.521810391,-0.313535314,0.408607177],[0,0,0,0],[9E+09,9E+09,9E+09,9E+09,9E+09,9E+09]];
    CONST robtarget Target_LetFron1_1310:=[[30.151,-121.309,47.417],[0.680036541,-0.521810391,-0.313535314,0.408607177],[0,0,0,0],[9E+09,9E+09,9E+09,9E+09,9E+09,9E+09]];
    CONST robtarget Target_LetFron1_1320:=[[29.67,-121.428,47.148],[0.680036541,-0.521810391,-0.313535314,0.408607177],[0,0,0,0],[9E+09,9E+09,9E+09,9E+09,9E+09,9E+09]];
    CONST robtarget Target_LetFron1_1330:=[[29.175,-121.548,46.863],[0.680036541,-0.521810391,-0.313535314,0.408607177],[0,0,0,0],[9E+09,9E+09,9E+09,9E+09,9E+09,9E+09]];
    CONST robtarget Target_LetFron1_1340:=[[28.372,-121.737,46.72],[0.680036541,-0.521810391,-0.313535314,0.408607177],[0,0,0,0],[9E+09,9E+09,9E+09,9E+09,9E+09,9E+09]];
    CONST robtarget Target_LetFron1_1350:=[[27.576,-121.92,46.773],[0.680036541,-0.521810391,-0.313535314,0.408607177],[0,0,0,0],[9E+09,9E+09,9E+09,9E+09,9E+09,9E+09]];
    CONST robtarget Target_LetFron1_1360:=[[37.518,-141.934,46.78],[0.680036541,-0.521810391,-0.313535314,0.408607177],[0,0,0,0],[9E+09,9E+09,9E+09,9E+09,9E+09,9E+09]];
    CONST robtarget Target_LetFron1_1370:=[[35.07,-142.46,57.11],[0.680036541,-0.521810391,-0.313535314,0.408607177],[0,0,0,0],[9E+09,9E+09,9E+09,9E+09,9E+09,9E+09]];
    CONST robtarget Target_LetFron1_1380:=[[25.07,-122.46,57.11],[0.680036541,-0.521810391,-0.313535314,0.408607177],[0,0,0,0],[9E+09,9E+09,9E+09,9E+09,9E+09,9E+09]];
    CONST robtarget Target_LetFron1_1390:=[[25.07,-122.46,46.866],[0.680036541,-0.521810391,-0.313535314,0.408607177],[0,0,0,0],[9E+09,9E+09,9E+09,9E+09,9E+09,9E+09]];
    CONST robtarget Target_LetFron1_1400:=[[35.07,-142.46,46.866],[0.680036541,-0.521810391,-0.313535314,0.408607177],[0,0,0,0],[9E+09,9E+09,9E+09,9E+09,9E+09,9E+09]];
    CONST robtarget Target_LetFron1_1410:=[[35.063,-142.462,44.786],[0.680036541,-0.521810391,-0.313535314,0.408607177],[0,0,0,0],[9E+09,9E+09,9E+09,9E+09,9E+09,9E+09]];
    CONST robtarget Target_LetFron1_1420:=[[25.063,-122.462,44.786],[0.680036541,-0.521810391,-0.313535314,0.408607177],[0,0,0,0],[9E+09,9E+09,9E+09,9E+09,9E+09,9E+09]];
    CONST robtarget Target_LetFron1_1430:=[[35.063,-142.462,44.786],[0.680036541,-0.521810391,-0.313535314,0.408607177],[0,0,0,0],[9E+09,9E+09,9E+09,9E+09,9E+09,9E+09]];
    CONST robtarget Target_LetFron1_1440:=[[29.75,-143.43,47.59],[0.680036541,-0.521810391,-0.313535314,0.408607177],[0,0,0,0],[9E+09,9E+09,9E+09,9E+09,9E+09,9E+09]];
    CONST robtarget Target_LetFron1_1450:=[[19.75,-123.43,47.59],[0.680036541,-0.521810391,-0.313535314,0.408607177],[0,0,0,0],[9E+09,9E+09,9E+09,9E+09,9E+09,9E+09]];
    CONST robtarget Target_LetFron1_1460:=[[20.377,-123.328,48.171],[0.680036541,-0.521810391,-0.313535314,0.408607177],[0,0,0,0],[9E+09,9E+09,9E+09,9E+09,9E+09,9E+09]];
    CONST robtarget Target_LetFron1_1470:=[[20.919,-123.237,48.849],[0.680036541,-0.521810391,-0.313535314,0.408607177],[0,0,0,0],[9E+09,9E+09,9E+09,9E+09,9E+09,9E+09]];
    CONST robtarget Target_LetFron1_1480:=[[21.332,-123.166,49.674],[0.680036541,-0.521810391,-0.313535314,0.408607177],[0,0,0,0],[9E+09,9E+09,9E+09,9E+09,9E+09,9E+09]];
    CONST robtarget Target_LetFron1_1490:=[[21.746,-123.094,51.083],[0.680036541,-0.521810391,-0.313535314,0.408607177],[0,0,0,0],[9E+09,9E+09,9E+09,9E+09,9E+09,9E+09]];
    CONST robtarget Target_LetFron1_1500:=[[21.746,-123.094,52.253],[0.680036541,-0.521810391,-0.313535314,0.408607177],[0,0,0,0],[9E+09,9E+09,9E+09,9E+09,9E+09,9E+09]];
    CONST robtarget Target_LetFron1_1510:=[[21.602,-123.119,53.771],[0.680036541,-0.521810391,-0.313535314,0.408607177],[0,0,0,0],[9E+09,9E+09,9E+09,9E+09,9E+09,9E+09]];
    CONST robtarget Target_LetFron1_1520:=[[21.362,-123.161,54.659],[0.680036541,-0.521810391,-0.313535314,0.408607177],[0,0,0,0],[9E+09,9E+09,9E+09,9E+09,9E+09,9E+09]];
    CONST robtarget Target_LetFron1_1530:=[[20.771,-123.262,55.806],[0.680036541,-0.521810391,-0.313535314,0.408607177],[0,0,0,0],[9E+09,9E+09,9E+09,9E+09,9E+09,9E+09]];
    CONST robtarget Target_LetFron1_1540:=[[19.905,-123.405,56.593],[0.680036541,-0.521810391,-0.313535314,0.408607177],[0,0,0,0],[9E+09,9E+09,9E+09,9E+09,9E+09,9E+09]];
    CONST robtarget Target_LetFron1_1550:=[[18.127,-123.679,57.403],[0.680036541,-0.521810391,-0.313535314,0.408607177],[0,0,0,0],[9E+09,9E+09,9E+09,9E+09,9E+09,9E+09]];
    CONST robtarget Target_LetFron1_1560:=[[16.241,-123.94,57.403],[0.680036541,-0.521810391,-0.313535314,0.408607177],[0,0,0,0],[9E+09,9E+09,9E+09,9E+09,9E+09,9E+09]];
    CONST robtarget Target_LetFron1_1570:=[[14.604,-124.144,56.751],[0.680036541,-0.521810391,-0.313535314,0.408607177],[0,0,0,0],[9E+09,9E+09,9E+09,9E+09,9E+09,9E+09]];
    CONST robtarget Target_LetFron1_1580:=[[13.599,-124.258,55.935],[0.680036541,-0.521810391,-0.313535314,0.408607177],[0,0,0,0],[9E+09,9E+09,9E+09,9E+09,9E+09,9E+09]];
    CONST robtarget Target_LetFron1_1590:=[[12.861,-124.337,54.839],[0.680036541,-0.521810391,-0.313535314,0.408607177],[0,0,0,0],[9E+09,9E+09,9E+09,9E+09,9E+09,9E+09]];
    CONST robtarget Target_LetFron1_1600:=[[12.234,-124.4,53.002],[0.680036541,-0.521810391,-0.313535314,0.408607177],[0,0,0,0],[9E+09,9E+09,9E+09,9E+09,9E+09,9E+09]];
    CONST robtarget Target_LetFron1_1610:=[[12.374,-124.386,50.335],[0.680036541,-0.521810391,-0.313535314,0.408607177],[0,0,0,0],[9E+09,9E+09,9E+09,9E+09,9E+09,9E+09]];
    CONST robtarget Target_LetFron1_1620:=[[12.98,-124.324,48.699],[0.680036541,-0.521810391,-0.313535314,0.408607177],[0,0,0,0],[9E+09,9E+09,9E+09,9E+09,9E+09,9E+09]];
    CONST robtarget Target_LetFron1_1630:=[[14.024,-124.211,47.53],[0.680036541,-0.521810391,-0.313535314,0.408607177],[0,0,0,0],[9E+09,9E+09,9E+09,9E+09,9E+09,9E+09]];
    CONST robtarget Target_LetFron1_1640:=[[15.431,-124.044,46.872],[0.680036541,-0.521810391,-0.313535314,0.408607177],[0,0,0,0],[9E+09,9E+09,9E+09,9E+09,9E+09,9E+09]];
    CONST robtarget Target_LetFron1_1650:=[[17.199,-123.811,46.72],[0.680036541,-0.521810391,-0.313535314,0.408607177],[0,0,0,0],[9E+09,9E+09,9E+09,9E+09,9E+09,9E+09]];
    CONST robtarget Target_LetFron1_1660:=[[18.168,-123.673,46.829],[0.680036541,-0.521810391,-0.313535314,0.408607177],[0,0,0,0],[9E+09,9E+09,9E+09,9E+09,9E+09,9E+09]];
    CONST robtarget Target_LetFron1_1670:=[[19.75,-123.43,47.59],[0.680036541,-0.521810391,-0.313535314,0.408607177],[0,0,0,0],[9E+09,9E+09,9E+09,9E+09,9E+09,9E+09]];
    CONST robtarget Target_LetFron1_1680:=[[29.75,-143.43,47.59],[0.680036541,-0.521810391,-0.313535314,0.408607177],[0,0,0,0],[9E+09,9E+09,9E+09,9E+09,9E+09,9E+09]];
    !***********************************************************
    !Dibujo segundo cuadrante de letrero frontal
    CONST robtarget Target_LetFron2_10:=[[19.88,-144.609,74.943],[0.680036541,-0.521810391,-0.313535314,0.408607177],[0,0,0,0],[9E+09,9E+09,9E+09,9E+09,9E+09,9E+09]];
    CONST robtarget Target_LetFron2_20:=[[9.88,-124.609,74.943],[0.680036541,-0.521810391,-0.313535314,0.408607177],[0,0,0,0],[9E+09,9E+09,9E+09,9E+09,9E+09,9E+09]];
    CONST robtarget Target_LetFron2_30:=[[11.251,-124.493,73.811],[0.680036541,-0.521810391,-0.313535314,0.408607177],[0,0,0,0],[9E+09,9E+09,9E+09,9E+09,9E+09,9E+09]];
    CONST robtarget Target_LetFron2_40:=[[12.534,-124.37,73.706],[0.680036541,-0.521810391,-0.313535314,0.408607177],[0,0,0,0],[9E+09,9E+09,9E+09,9E+09,9E+09,9E+09]];
    CONST robtarget Target_LetFron2_50:=[[14.383,-124.17,73.976],[0.680036541,-0.521810391,-0.313535314,0.408607177],[0,0,0,0],[9E+09,9E+09,9E+09,9E+09,9E+09,9E+09]];
    CONST robtarget Target_LetFron2_60:=[[15.432,-124.044,74.542],[0.680036541,-0.521810391,-0.313535314,0.408607177],[0,0,0,0],[9E+09,9E+09,9E+09,9E+09,9E+09,9E+09]];
    CONST robtarget Target_LetFron2_70:=[[15.826,-123.994,74.943],[0.680036541,-0.521810391,-0.313535314,0.408607177],[0,0,0,0],[9E+09,9E+09,9E+09,9E+09,9E+09,9E+09]];
    CONST robtarget Target_LetFron2_80:=[[16.325,-123.929,75.618],[0.680036541,-0.521810391,-0.313535314,0.408607177],[0,0,0,0],[9E+09,9E+09,9E+09,9E+09,9E+09,9E+09]];
    CONST robtarget Target_LetFron2_90:=[[16.488,-123.908,76.675],[0.680036541,-0.521810391,-0.313535314,0.408607177],[0,0,0,0],[9E+09,9E+09,9E+09,9E+09,9E+09,9E+09]];
    CONST robtarget Target_LetFron2_100:=[[16.384,-123.922,77.642],[0.680036541,-0.521810391,-0.313535314,0.408607177],[0,0,0,0],[9E+09,9E+09,9E+09,9E+09,9E+09,9E+09]];
    CONST robtarget Target_LetFron2_110:=[[15.802,-123.997,78.469],[0.680036541,-0.521810391,-0.313535314,0.408607177],[0,0,0,0],[9E+09,9E+09,9E+09,9E+09,9E+09,9E+09]];
    CONST robtarget Target_LetFron2_120:=[[15.187,-124.074,78.939],[0.680036541,-0.521810391,-0.313535314,0.408607177],[0,0,0,0],[9E+09,9E+09,9E+09,9E+09,9E+09,9E+09]];
    CONST robtarget Target_LetFron2_160:=[[14.346,-124.174,79.351],[0.680036541,-0.521810391,-0.313535314,0.408607177],[0,0,0,0],[9E+09,9E+09,9E+09,9E+09,9E+09,9E+09]];
    CONST robtarget Target_LetFron2_200:=[[13.608,-124.257,79.644],[0.680036541,-0.521810391,-0.313535314,0.408607177],[0,0,0,0],[9E+09,9E+09,9E+09,9E+09,9E+09,9E+09]];
    CONST robtarget Target_LetFron2_210:=[[12.736,-124.35,79.989],[0.680036541,-0.521810391,-0.313535314,0.408607177],[0,0,0,0],[9E+09,9E+09,9E+09,9E+09,9E+09,9E+09]];
    CONST robtarget Target_LetFron2_220:=[[11.796,-124.442,80.513],[0.680036541,-0.521810391,-0.313535314,0.408607177],[0,0,0,0],[9E+09,9E+09,9E+09,9E+09,9E+09,9E+09]];
    CONST robtarget Target_LetFron2_230:=[[9.51,-124.638,81.195],[0.680036541,-0.521810391,-0.313535314,0.408607177],[0,0,0,0],[9E+09,9E+09,9E+09,9E+09,9E+09,9E+09]];
    CONST robtarget Target_LetFron2_250:=[[9.682,-124.624,82.38],[0.680036541,-0.521810391,-0.313535314,0.408607177],[0,0,0,0],[9E+09,9E+09,9E+09,9E+09,9E+09,9E+09]];
    CONST robtarget Target_LetFron2_260:=[[10.026,-124.597,82.86],[0.680036541,-0.521810391,-0.313535314,0.408607177],[0,0,0,0],[9E+09,9E+09,9E+09,9E+09,9E+09,9E+09]];
    CONST robtarget Target_LetFron2_270:=[[10.848,-124.528,83.714],[0.680036541,-0.521810391,-0.313535314,0.408607177],[0,0,0,0],[9E+09,9E+09,9E+09,9E+09,9E+09,9E+09]];
    CONST robtarget Target_LetFron2_280:=[[11.759,-124.446,84.119],[0.680036541,-0.521810391,-0.313535314,0.408607177],[0,0,0,0],[9E+09,9E+09,9E+09,9E+09,9E+09,9E+09]];
    CONST robtarget Target_LetFron2_290:=[[12.743,-124.349,84.389],[0.680036541,-0.521810391,-0.313535314,0.408607177],[0,0,0,0],[9E+09,9E+09,9E+09,9E+09,9E+09,9E+09]];
    CONST robtarget Target_LetFron2_300:=[[13.832,-124.232,84.389],[0.680036541,-0.521810391,-0.313535314,0.408607177],[0,0,0,0],[9E+09,9E+09,9E+09,9E+09,9E+09,9E+09]];
    CONST robtarget Target_LetFron2_310:=[[14.446,-124.162,84.355],[0.680036541,-0.521810391,-0.313535314,0.408607177],[0,0,0,0],[9E+09,9E+09,9E+09,9E+09,9E+09,9E+09]];
    CONST robtarget Target_LetFron2_320:=[[15.038,-124.092,84.254],[0.680036541,-0.521810391,-0.313535314,0.408607177],[0,0,0,0],[9E+09,9E+09,9E+09,9E+09,9E+09,9E+09]];
    CONST robtarget Target_LetFron2_330:=[[16.566,-123.897,83.04],[0.680036541,-0.521810391,-0.313535314,0.408607177],[0,0,0,0],[9E+09,9E+09,9E+09,9E+09,9E+09,9E+09]];
    CONST robtarget Target_LetFron2_340:=[[26.566,-143.897,83.04],[0.680036541,-0.521810391,-0.313535314,0.408607177],[0,0,0,0],[9E+09,9E+09,9E+09,9E+09,9E+09,9E+09]];
    CONST robtarget Target_LetFron2_350:=[[28.695,-143.594,83.699],[0.680036541,-0.521810391,-0.313535314,0.408607177],[0,0,0,0],[9E+09,9E+09,9E+09,9E+09,9E+09,9E+09]];
    CONST robtarget Target_LetFron2_360:=[[18.695,-123.594,83.699],[0.680036541,-0.521810391,-0.313535314,0.408607177],[0,0,0,0],[9E+09,9E+09,9E+09,9E+09,9E+09,9E+09]];
    CONST robtarget Target_LetFron2_370:=[[19.54,-123.463,84.014],[0.680036541,-0.521810391,-0.313535314,0.408607177],[0,0,0,0],[9E+09,9E+09,9E+09,9E+09,9E+09,9E+09]];
    CONST robtarget Target_LetFron2_380:=[[20.465,-123.313,84.239],[0.680036541,-0.521810391,-0.313535314,0.408607177],[0,0,0,0],[9E+09,9E+09,9E+09,9E+09,9E+09,9E+09]];
    CONST robtarget Target_LetFron2_390:=[[22.046,-123.041,84.389],[0.680036541,-0.521810391,-0.313535314,0.408607177],[0,0,0,0],[9E+09,9E+09,9E+09,9E+09,9E+09,9E+09]];
    CONST robtarget Target_LetFron2_400:=[[23.682,-122.736,84.209],[0.680036541,-0.521810391,-0.313535314,0.408607177],[0,0,0,0],[9E+09,9E+09,9E+09,9E+09,9E+09,9E+09]];
    CONST robtarget Target_LetFron2_410:=[[25.079,-122.458,83.489],[0.680036541,-0.521810391,-0.313535314,0.408607177],[0,0,0,0],[9E+09,9E+09,9E+09,9E+09,9E+09,9E+09]];
    CONST robtarget Target_LetFron2_420:=[[25.637,-122.343,82.935],[0.680036541,-0.521810391,-0.313535314,0.408607177],[0,0,0,0],[9E+09,9E+09,9E+09,9E+09,9E+09,9E+09]];
    CONST robtarget Target_LetFron2_430:=[[26.575,-122.142,80.937],[0.680036541,-0.521810391,-0.313535314,0.408607177],[0,0,0,0],[9E+09,9E+09,9E+09,9E+09,9E+09,9E+09]];
    CONST robtarget Target_LetFron2_440:=[[26.678,-122.12,79.869],[0.680036541,-0.521810391,-0.313535314,0.408607177],[0,0,0,0],[9E+09,9E+09,9E+09,9E+09,9E+09,9E+09]];
    CONST robtarget Target_LetFron2_450:=[[26.535,-122.151,77.625],[0.680036541,-0.521810391,-0.313535314,0.408607177],[0,0,0,0],[9E+09,9E+09,9E+09,9E+09,9E+09,9E+09]];
    CONST robtarget Target_LetFron2_460:=[[25.908,-122.286,75.828],[0.680036541,-0.521810391,-0.313535314,0.408607177],[0,0,0,0],[9E+09,9E+09,9E+09,9E+09,9E+09,9E+09]];
    CONST robtarget Target_LetFron2_470:=[[24.476,-122.58,74.359],[0.680036541,-0.521810391,-0.313535314,0.408607177],[0,0,0,0],[9E+09,9E+09,9E+09,9E+09,9E+09,9E+09]];
    CONST robtarget Target_LetFron2_480:=[[23.367,-122.797,73.87],[0.680036541,-0.521810391,-0.313535314,0.408607177],[0,0,0,0],[9E+09,9E+09,9E+09,9E+09,9E+09,9E+09]];
    CONST robtarget Target_LetFron2_490:=[[21.81,-123.083,73.706],[0.680036541,-0.521810391,-0.313535314,0.408607177],[0,0,0,0],[9E+09,9E+09,9E+09,9E+09,9E+09,9E+09]];
    CONST robtarget Target_LetFron2_500:=[[20.539,-123.301,73.999],[0.680036541,-0.521810391,-0.313535314,0.408607177],[0,0,0,0],[9E+09,9E+09,9E+09,9E+09,9E+09,9E+09]];
    CONST robtarget Target_LetFron2_510:=[[19.555,-123.461,74.636],[0.680036541,-0.521810391,-0.313535314,0.408607177],[0,0,0,0],[9E+09,9E+09,9E+09,9E+09,9E+09,9E+09]];
    CONST robtarget Target_LetFron2_520:=[[18.866,-123.568,75.543],[0.680036541,-0.521810391,-0.313535314,0.408607177],[0,0,0,0],[9E+09,9E+09,9E+09,9E+09,9E+09,9E+09]];
    CONST robtarget Target_LetFron2_530:=[[18.717,-123.591,76.023],[0.680036541,-0.521810391,-0.313535314,0.408607177],[0,0,0,0],[9E+09,9E+09,9E+09,9E+09,9E+09,9E+09]];
    CONST robtarget Target_LetFron2_540:=[[18.473,-123.627,76.997],[0.680036541,-0.521810391,-0.313535314,0.408607177],[0,0,0,0],[9E+09,9E+09,9E+09,9E+09,9E+09,9E+09]];
    CONST robtarget Target_LetFron2_550:=[[18.48,-123.626,78.017],[0.680036541,-0.521810391,-0.313535314,0.408607177],[0,0,0,0],[9E+09,9E+09,9E+09,9E+09,9E+09,9E+09]];
    CONST robtarget Target_LetFron2_560:=[[18.54,-123.617,78.857],[0.680036541,-0.521810391,-0.313535314,0.408607177],[0,0,0,0],[9E+09,9E+09,9E+09,9E+09,9E+09,9E+09]];
    CONST robtarget Target_LetFron2_570:=[[21.669,-123.107,78.857],[0.680036541,-0.521810391,-0.313535314,0.408607177],[0,0,0,0],[9E+09,9E+09,9E+09,9E+09,9E+09,9E+09]];
    CONST robtarget Target_LetFron2_580:=[[24.785,-122.518,78.857],[0.680036541,-0.521810391,-0.313535314,0.408607177],[0,0,0,0],[9E+09,9E+09,9E+09,9E+09,9E+09,9E+09]];
    CONST robtarget Target_LetFron2_590:=[[34.785,-142.518,78.857],[0.680036541,-0.521810391,-0.313535314,0.408607177],[0,0,0,0],[9E+09,9E+09,9E+09,9E+09,9E+09,9E+09]];
    CONST robtarget Target_LetFron2_600:=[[37.559,-141.924,83.782],[0.680036541,-0.521810391,-0.313535314,0.408607177],[0,0,0,0],[9E+09,9E+09,9E+09,9E+09,9E+09,9E+09]];
    CONST robtarget Target_LetFron2_610:=[[27.559,-121.924,83.782],[0.680036541,-0.521810391,-0.313535314,0.408607177],[0,0,0,0],[9E+09,9E+09,9E+09,9E+09,9E+09,9E+09]];
    CONST robtarget Target_LetFron2_620:=[[29.274,-121.524,84.337],[0.680036541,-0.521810391,-0.313535314,0.408607177],[0,0,0,0],[9E+09,9E+09,9E+09,9E+09,9E+09,9E+09]];
    CONST robtarget Target_LetFron2_630:=[[30.671,-121.179,84.389],[0.680036541,-0.521810391,-0.313535314,0.408607177],[0,0,0,0],[9E+09,9E+09,9E+09,9E+09,9E+09,9E+09]];
    CONST robtarget Target_LetFron2_640:=[[31.746,-120.902,83.999],[0.680036541,-0.521810391,-0.313535314,0.408607177],[0,0,0,0],[9E+09,9E+09,9E+09,9E+09,9E+09,9E+09]];
    CONST robtarget Target_LetFron2_650:=[[32.535,-120.692,83.242],[0.680036541,-0.521810391,-0.313535314,0.408607177],[0,0,0,0],[9E+09,9E+09,9E+09,9E+09,9E+09,9E+09]];
    CONST robtarget Target_LetFron2_660:=[[32.883,-120.597,82.058],[0.680036541,-0.521810391,-0.313535314,0.408607177],[0,0,0,0],[9E+09,9E+09,9E+09,9E+09,9E+09,9E+09]];
    CONST robtarget Target_LetFron2_670:=[[32.774,-120.627,72.267],[0.680036541,-0.521810391,-0.313535314,0.408607177],[0,0,0,0],[9E+09,9E+09,9E+09,9E+09,9E+09,9E+09]];
    CONST robtarget Target_LetFron2_680:=[[32.796,-120.621,73.976],[0.680036541,-0.521810391,-0.313535314,0.408607177],[0,0,0,0],[9E+09,9E+09,9E+09,9E+09,9E+09,9E+09]];
    CONST robtarget Target_LetFron2_690:=[[34.421,-120.167,74.201],[0.680036541,-0.521810391,-0.313535314,0.408607177],[0,0,0,0],[9E+09,9E+09,9E+09,9E+09,9E+09,9E+09]];
    CONST robtarget Target_LetFron2_700:=[[27.756,-121.879,73.976],[0.680036541,-0.521810391,-0.313535314,0.408607177],[0,0,0,0],[9E+09,9E+09,9E+09,9E+09,9E+09,9E+09]];
    CONST robtarget Target_LetFron2_710:=[[37.756,-141.879,73.976],[0.680036541,-0.521810391,-0.313535314,0.408607177],[0,0,0,0],[9E+09,9E+09,9E+09,9E+09,9E+09,9E+09]];
    CONST robtarget Target_LetFron2_720:=[[46.102,-129.673,84.097],[0.680036541,-0.521810391,-0.313535314,0.408607177],[0,0,0,0],[9E+09,9E+09,9E+09,9E+09,9E+09,9E+09]];
    CONST robtarget Target_LetFron2_730:=[[36.102,-119.673,84.097],[0.680036541,-0.521810391,-0.313535314,0.408607177],[0,0,0,0],[9E+09,9E+09,9E+09,9E+09,9E+09,9E+09]];
    CONST robtarget Target_LetFron2_740:=[[36.102,-119.673,76.083],[0.680036541,-0.521810391,-0.313535314,0.408607177],[0,0,0,0],[9E+09,9E+09,9E+09,9E+09,9E+09,9E+09]];
    CONST robtarget Target_LetFron2_750:=[[36.59,-119.525,74.876],[0.680036541,-0.521810391,-0.313535314,0.408607177],[0,0,0,0],[9E+09,9E+09,9E+09,9E+09,9E+09,9E+09]];
    CONST robtarget Target_LetFron2_760:=[[37.278,-119.312,74.186],[0.680036541,-0.521810391,-0.313535314,0.408607177],[0,0,0,0],[9E+09,9E+09,9E+09,9E+09,9E+09,9E+09]];
    CONST robtarget Target_LetFron2_770:=[[38.203,-119.019,73.766],[0.680036541,-0.521810391,-0.313535314,0.408607177],[0,0,0,0],[9E+09,9E+09,9E+09,9E+09,9E+09,9E+09]];
    CONST robtarget Target_LetFron2_780:=[[39.062,-118.74,73.706],[0.680036541,-0.521810391,-0.313535314,0.408607177],[0,0,0,0],[9E+09,9E+09,9E+09,9E+09,9E+09,9E+09]];
    CONST robtarget Target_LetFron2_790:=[[39.745,-118.513,73.766],[0.680036541,-0.521810391,-0.313535314,0.408607177],[0,0,0,0],[9E+09,9E+09,9E+09,9E+09,9E+09,9E+09]];
    CONST robtarget Target_LetFron2_800:=[[40.512,-118.253,74.006],[0.680036541,-0.521810391,-0.313535314,0.408607177],[0,0,0,0],[9E+09,9E+09,9E+09,9E+09,9E+09,9E+09]];
    CONST robtarget Target_LetFron2_810:=[[41.624,-117.866,74.501],[0.680036541,-0.521810391,-0.313535314,0.408607177],[0,0,0,0],[9E+09,9E+09,9E+09,9E+09,9E+09,9E+09]];
    CONST robtarget Target_LetFron2_820:=[[42.09,-117.701,74.748],[0.680036541,-0.521810391,-0.313535314,0.408607177],[0,0,0,0],[9E+09,9E+09,9E+09,9E+09,9E+09,9E+09]];
    CONST robtarget Target_LetFron2_830:=[[42.57,-117.528,73.706],[0.680036541,-0.521810391,-0.313535314,0.408607177],[0,0,0,0],[9E+09,9E+09,9E+09,9E+09,9E+09,9E+09]];
    CONST robtarget Target_LetFron2_840:=[[43.224,-117.289,73.853],[0.680036541,-0.521810391,-0.313535314,0.408607177],[0,0,0,0],[9E+09,9E+09,9E+09,9E+09,9E+09,9E+09]];
    CONST robtarget Target_LetFron2_850:=[[42.971,-117.382,84.097],[0.680036541,-0.521810391,-0.313535314,0.408607177],[0,0,0,0],[9E+09,9E+09,9E+09,9E+09,9E+09,9E+09]];
    CONST robtarget Target_LetFron2_860:=[[52.971,-127.382,84.097],[0.680036541,-0.521810391,-0.313535314,0.408607177],[0,0,0,0],[9E+09,9E+09,9E+09,9E+09,9E+09,9E+09]];
    CONST robtarget Target_LetFron2_870:=[[56.087,-136.194,83.579],[0.680036541,-0.521810391,-0.313535314,0.408607177],[0,0,0,0],[9E+09,9E+09,9E+09,9E+09,9E+09,9E+09]];
    CONST robtarget Target_LetFron2_880:=[[46.087,-116.194,83.579],[0.680036541,-0.521810391,-0.313535314,0.408607177],[0,0,0,0],[9E+09,9E+09,9E+09,9E+09,9E+09,9E+09]];
    CONST robtarget Target_LetFron2_890:=[[47.422,-115.655,84.089],[0.680036541,-0.521810391,-0.313535314,0.408607177],[0,0,0,0],[9E+09,9E+09,9E+09,9E+09,9E+09,9E+09]];
    CONST robtarget Target_LetFron2_900:=[[48.58,-115.174,84.333],[0.680036541,-0.521810391,-0.313535314,0.408607177],[0,0,0,0],[9E+09,9E+09,9E+09,9E+09,9E+09,9E+09]];
    CONST robtarget Target_LetFron2_910:=[[50.618,-114.293,84.254],[0.680036541,-0.521810391,-0.313535314,0.408607177],[0,0,0,0],[9E+09,9E+09,9E+09,9E+09,9E+09,9E+09]];
    CONST robtarget Target_LetFron2_920:=[[52.295,-113.535,83.489],[0.680036541,-0.521810391,-0.313535314,0.408607177],[0,0,0,0],[9E+09,9E+09,9E+09,9E+09,9E+09,9E+09]];
    CONST robtarget Target_LetFron2_930:=[[0.104,125,4.999],[0.680036541,-0.521810391,-0.313535314,0.408607177],[0,0,0,0],[9E+09,9E+09,9E+09,9E+09,9E+09,9E+09]];
    CONST robtarget Target_LetFron2_940:=[[53.206,-113.111,82.185],[0.680036541,-0.521810391,-0.313535314,0.408607177],[0,0,0,0],[9E+09,9E+09,9E+09,9E+09,9E+09,9E+09]];
    CONST robtarget Target_LetFron2_950:=[[53.775,-112.842,80.453],[0.680036541,-0.521810391,-0.313535314,0.408607177],[0,0,0,0],[9E+09,9E+09,9E+09,9E+09,9E+09,9E+09]];
    CONST robtarget Target_LetFron2_960:=[[53.775,-112.842,78.684],[0.680036541,-0.521810391,-0.313535314,0.408607177],[0,0,0,0],[9E+09,9E+09,9E+09,9E+09,9E+09,9E+09]];
    CONST robtarget Target_LetFron2_970:=[[53.687,-112.884,77.578],[0.680036541,-0.521810391,-0.313535314,0.408607177],[0,0,0,0],[9E+09,9E+09,9E+09,9E+09,9E+09,9E+09]];
    CONST robtarget Target_LetFron2_980:=[[52.88,-113.264,75.408],[0.680036541,-0.521810391,-0.313535314,0.408607177],[0,0,0,0],[9E+09,9E+09,9E+09,9E+09,9E+09,9E+09]];
    CONST robtarget Target_LetFron2_990:=[[52.057,-113.645,74.569],[0.680036541,-0.521810391,-0.313535314,0.408607177],[0,0,0,0],[9E+09,9E+09,9E+09,9E+09,9E+09,9E+09]];
    CONST robtarget Target_LetFron2_1000:=[[51.094,-114.081,73.924],[0.680036541,-0.521810391,-0.313535314,0.408607177],[0,0,0,0],[9E+09,9E+09,9E+09,9E+09,9E+09,9E+09]];
    CONST robtarget Target_LetFron2_1010:=[[49.949,-114.587,73.706],[0.680036541,-0.521810391,-0.313535314,0.408607177],[0,0,0,0],[9E+09,9E+09,9E+09,9E+09,9E+09,9E+09]];
    CONST robtarget Target_LetFron2_1020:=[[48.274,-115.302,73.901],[0.680036541,-0.521810391,-0.313535314,0.408607177],[0,0,0,0],[9E+09,9E+09,9E+09,9E+09,9E+09,9E+09]];
    CONST robtarget Target_LetFron2_1030:=[[47.144,-115.769,74.636],[0.680036541,-0.521810391,-0.313535314,0.408607177],[0,0,0,0],[9E+09,9E+09,9E+09,9E+09,9E+09,9E+09]];
    CONST robtarget Target_LetFron2_1040:=[[46.282,-116.116,76.255],[0.680036541,-0.521810391,-0.313535314,0.408607177],[0,0,0,0],[9E+09,9E+09,9E+09,9E+09,9E+09,9E+09]];
    CONST robtarget Target_LetFron2_1050:=[[46.129,-116.177,77.777],[0.680036541,-0.521810391,-0.313535314,0.408607177],[0,0,0,0],[9E+09,9E+09,9E+09,9E+09,9E+09,9E+09]];
    CONST robtarget Target_LetFron2_1060:=[[46.191,-116.152,78.857],[0.680036541,-0.521810391,-0.313535314,0.408607177],[0,0,0,0],[9E+09,9E+09,9E+09,9E+09,9E+09,9E+09]];
    CONST robtarget Target_LetFron2_1070:=[[49.123,-114.943,78.857],[0.680036541,-0.521810391,-0.313535314,0.408607177],[0,0,0,0],[9E+09,9E+09,9E+09,9E+09,9E+09,9E+09]];
    CONST robtarget Target_LetFron2_1080:=[[52.023,-113.66,78.857],[0.680036541,-0.521810391,-0.313535314,0.408607177],[0,0,0,0],[9E+09,9E+09,9E+09,9E+09,9E+09,9E+09]];
    CONST robtarget Target_LetFron2_1090:=[[62.023,-133.66,78.857],[0.680036541,-0.521810391,-0.313535314,0.408607177],[0,0,0,0],[9E+09,9E+09,9E+09,9E+09,9E+09,9E+09]];
    CONST robtarget Target_LetFron2_1100:=[[70.754,-129.243,83.489],[0.680036541,-0.521810391,-0.313535314,0.408607177],[0,0,0,0],[9E+09,9E+09,9E+09,9E+09,9E+09,9E+09]];
    CONST robtarget Target_LetFron2_1110:=[[60.754,-109.243,83.489],[0.680036541,-0.521810391,-0.313535314,0.408607177],[0,0,0,0],[9E+09,9E+09,9E+09,9E+09,9E+09,9E+09]];
    CONST robtarget Target_LetFron2_1120:=[[61.929,-108.581,84.389],[0.680036541,-0.521810391,-0.313535314,0.408607177],[0,0,0,0],[9E+09,9E+09,9E+09,9E+09,9E+09,9E+09]];
    CONST robtarget Target_LetFron2_1130:=[[63.079,-107.917,86.391],[0.680036541,-0.521810391,-0.313535314,0.408607177],[0,0,0,0],[9E+09,9E+09,9E+09,9E+09,9E+09,9E+09]];
    CONST robtarget Target_LetFron2_1140:=[[62.69,-108.143,87.65],[0.680036541,-0.521810391,-0.313535314,0.408607177],[0,0,0,0],[9E+09,9E+09,9E+09,9E+09,9E+09,9E+09]];
    CONST robtarget Target_LetFron2_1150:=[[60.773,-109.232,88.701],[0.680036541,-0.521810391,-0.313535314,0.408607177],[0,0,0,0],[9E+09,9E+09,9E+09,9E+09,9E+09,9E+09]];
    CONST robtarget Target_LetFron2_1160:=[[57.504,-110.988,88.235],[0.680036541,-0.521810391,-0.313535314,0.408607177],[0,0,0,0],[9E+09,9E+09,9E+09,9E+09,9E+09,9E+09]];
    CONST robtarget Target_LetFron2_1170:=[[56.529,-111.488,87.599],[0.680036541,-0.521810391,-0.313535314,0.408607177],[0,0,0,0],[9E+09,9E+09,9E+09,9E+09,9E+09,9E+09]];
    CONST robtarget Target_LetFron2_1180:=[[55.246,-112.129,85.828],[0.680036541,-0.521810391,-0.313535314,0.408607177],[0,0,0,0],[9E+09,9E+09,9E+09,9E+09,9E+09,9E+09]];
    CONST robtarget Target_LetFron2_1190:=[[55.075,-112.213,84.411],[0.680036541,-0.521810391,-0.313535314,0.408607177],[0,0,0,0],[9E+09,9E+09,9E+09,9E+09,9E+09,9E+09]];
    CONST robtarget Target_LetFron2_1200:=[[55.659,-111.924,83.175],[0.680036541,-0.521810391,-0.313535314,0.408607177],[0,0,0,0],[9E+09,9E+09,9E+09,9E+09,9E+09,9E+09]];
    CONST robtarget Target_LetFron2_1210:=[[56.824,-111.337,82.612],[0.680036541,-0.521810391,-0.313535314,0.408607177],[0,0,0,0],[9E+09,9E+09,9E+09,9E+09,9E+09,9E+09]];
    CONST robtarget Target_LetFron2_1220:=[[58.023,-110.717,82.41],[0.680036541,-0.521810391,-0.313535314,0.408607177],[0,0,0,0],[9E+09,9E+09,9E+09,9E+09,9E+09,9E+09]];
    CONST robtarget Target_LetFron2_1230:=[[60.065,-109.623,81.833],[0.680036541,-0.521810391,-0.313535314,0.408607177],[0,0,0,0],[9E+09,9E+09,9E+09,9E+09,9E+09,9E+09]];
    CONST robtarget Target_LetFron2_1240:=[[60.065,-109.623,80.881],[0.680036541,-0.521810391,-0.313535314,0.408607177],[0,0,0,0],[9E+09,9E+09,9E+09,9E+09,9E+09,9E+09]];
    CONST robtarget Target_LetFron2_1250:=[[59.215,-110.085,80.423],[0.680036541,-0.521810391,-0.313535314,0.408607177],[0,0,0,0],[9E+09,9E+09,9E+09,9E+09,9E+09,9E+09]];
    CONST robtarget Target_LetFron2_1260:=[[57.983,-110.738,80.161],[0.680036541,-0.521810391,-0.313535314,0.408607177],[0,0,0,0],[9E+09,9E+09,9E+09,9E+09,9E+09,9E+09]];
    CONST robtarget Target_LetFron2_1270:=[[56.579,-111.462,78.75],[0.680036541,-0.521810391,-0.313535314,0.408607177],[0,0,0,0],[9E+09,9E+09,9E+09,9E+09,9E+09,9E+09]];
    CONST robtarget Target_LetFron2_1280:=[[56.109,-111.7,77.17],[0.680036541,-0.521810391,-0.313535314,0.408607177],[0,0,0,0],[9E+09,9E+09,9E+09,9E+09,9E+09,9E+09]];
    CONST robtarget Target_LetFron2_1290:=[[56.323,-111.592,75.535],[0.680036541,-0.521810391,-0.313535314,0.408607177],[0,0,0,0],[9E+09,9E+09,9E+09,9E+09,9E+09,9E+09]];
    CONST robtarget Target_LetFron2_1300:=[[54.65,-112.42,75.393],[0.680036541,-0.521810391,-0.313535314,0.408607177],[0,0,0,0],[9E+09,9E+09,9E+09,9E+09,9E+09,9E+09]];
    CONST robtarget Target_LetFron2_1310:=[[54.65,-112.42,73.706],[0.680036541,-0.521810391,-0.313535314,0.408607177],[0,0,0,0],[9E+09,9E+09,9E+09,9E+09,9E+09,9E+09]];
    CONST robtarget Target_LetFron2_1320:=[[57.245,-111.122,74.269],[0.680036541,-0.521810391,-0.313535314,0.408607177],[0,0,0,0],[9E+09,9E+09,9E+09,9E+09,9E+09,9E+09]];
    CONST robtarget Target_LetFron2_1330:=[[58.719,-110.35,73.706],[0.680036541,-0.521810391,-0.313535314,0.408607177],[0,0,0,0],[9E+09,9E+09,9E+09,9E+09,9E+09,9E+09]];
    CONST robtarget Target_LetFron2_1340:=[[60.104,-109.602,73.813],[0.680036541,-0.521810391,-0.313535314,0.408607177],[0,0,0,0],[9E+09,9E+09,9E+09,9E+09,9E+09,9E+09]];
    CONST robtarget Target_LetFron2_1350:=[[61.284,-108.946,74.276],[0.680036541,-0.521810391,-0.313535314,0.408607177],[0,0,0,0],[9E+09,9E+09,9E+09,9E+09,9E+09,9E+09]];
    CONST robtarget Target_LetFron2_1360:=[[61.988,-108.547,74.831],[0.680036541,-0.521810391,-0.313535314,0.408607177],[0,0,0,0],[9E+09,9E+09,9E+09,9E+09,9E+09,9E+09]];
    CONST robtarget Target_LetFron2_1370:=[[62.45,-108.282,75.633],[0.680036541,-0.521810391,-0.313535314,0.408607177],[0,0,0,0],[9E+09,9E+09,9E+09,9E+09,9E+09,9E+09]];
    CONST robtarget Target_LetFron2_1380:=[[62.748,-108.11,76.907],[0.680036541,-0.521810391,-0.313535314,0.408607177],[0,0,0,0],[9E+09,9E+09,9E+09,9E+09,9E+09,9E+09]];
    CONST robtarget Target_LetFron2_1390:=[[62.607,-108.191,78.334],[0.680036541,-0.521810391,-0.313535314,0.408607177],[0,0,0,0],[9E+09,9E+09,9E+09,9E+09,9E+09,9E+09]];
    CONST robtarget Target_LetFron2_1400:=[[62.183,-108.435,79.194],[0.680036541,-0.521810391,-0.313535314,0.408607177],[0,0,0,0],[9E+09,9E+09,9E+09,9E+09,9E+09,9E+09]];
    CONST robtarget Target_LetFron2_1410:=[[61.329,-108.921,80.048],[0.680036541,-0.521810391,-0.313535314,0.408607177],[0,0,0,0],[9E+09,9E+09,9E+09,9E+09,9E+09,9E+09]];
    CONST robtarget Target_LetFron2_1420:=[[60.754,-109.243,80.228],[0.680036541,-0.521810391,-0.313535314,0.408607177],[0,0,0,0],[9E+09,9E+09,9E+09,9E+09,9E+09,9E+09]];
    CONST robtarget Target_LetFron2_1430:=[[70.754,-129.243,80.228],[0.680036541,-0.521810391,-0.313535314,0.408607177],[0,0,0,0],[9E+09,9E+09,9E+09,9E+09,9E+09,9E+09]];
    CONST robtarget Target_LetFron2_1440:=[[75.691,-126.347,84.097],[0.680036541,-0.521810391,-0.313535314,0.408607177],[0,0,0,0],[9E+09,9E+09,9E+09,9E+09,9E+09,9E+09]];
    CONST robtarget Target_LetFron2_1450:=[[65.691,-106.347,84.097],[0.680036541,-0.521810391,-0.313535314,0.408607177],[0,0,0,0],[9E+09,9E+09,9E+09,9E+09,9E+09,9E+09]];
    CONST robtarget Target_LetFron2_1460:=[[65.691,-106.347,73.853],[0.680036541,-0.521810391,-0.313535314,0.408607177],[0,0,0,0],[9E+09,9E+09,9E+09,9E+09,9E+09,9E+09]];
    CONST robtarget Target_LetFron2_1470:=[[75.691,-126.347,73.853],[0.680036541,-0.521810391,-0.313535314,0.408607177],[0,0,0,0],[9E+09,9E+09,9E+09,9E+09,9E+09,9E+09]];
    CONST robtarget Target_LetFron2_1480:=[[75.754,-126.308,69.298],[0.680036541,-0.521810391,-0.313535314,0.408607177],[0,0,0,0],[9E+09,9E+09,9E+09,9E+09,9E+09,9E+09]];
    CONST robtarget Target_LetFron2_1490:=[[65.799,-106.28,69.298],[0.680036541,-0.521810391,-0.313535314,0.408607177],[0,0,0,0],[9E+09,9E+09,9E+09,9E+09,9E+09,9E+09]];
    CONST robtarget Target_LetFron2_1500:=[[75.665,-126.363,69.298],[0.680036541,-0.521810391,-0.313535314,0.408607177],[0,0,0,0],[9E+09,9E+09,9E+09,9E+09,9E+09,9E+09]];
    CONST robtarget Target_LetFron2_1510:=[[78.402,-124.624,83.399],[0.680036541,-0.521810391,-0.313535314,0.408607177],[0,0,0,0],[9E+09,9E+09,9E+09,9E+09,9E+09,9E+09]];
    CONST robtarget Target_LetFron2_1520:=[[68.402,-104.624,83.399],[0.680036541,-0.521810391,-0.313535314,0.408607177],[0,0,0,0],[9E+09,9E+09,9E+09,9E+09,9E+09,9E+09]];
    CONST robtarget Target_LetFron2_1530:=[[71.196,-102.743,83.281],[0.680036541,-0.521810391,-0.313535314,0.408607177],[0,0,0,0],[9E+09,9E+09,9E+09,9E+09,9E+09,9E+09]];
    CONST robtarget Target_LetFron2_1540:=[[71.311,-102.663,68.916],[0.680036541,-0.521810391,-0.313535314,0.408607177],[0,0,0,0],[9E+09,9E+09,9E+09,9E+09,9E+09,9E+09]];
    CONST robtarget Target_LetFron2_1550:=[[81.311,-122.663,68.916],[0.680036541,-0.521810391,-0.313535314,0.408607177],[0,0,0,0],[9E+09,9E+09,9E+09,9E+09,9E+09,9E+09]];
    CONST robtarget Target_LetFron2_1560:=[[83.19,-121.333,83.579],[0.680036541,-0.521810391,-0.313535314,0.408607177],[0,0,0,0],[9E+09,9E+09,9E+09,9E+09,9E+09,9E+09]];
    CONST robtarget Target_LetFron2_1570:=[[73.19,-101.333,83.579],[0.680036541,-0.521810391,-0.313535314,0.408607177],[0,0,0,0],[9E+09,9E+09,9E+09,9E+09,9E+09,9E+09]];
    CONST robtarget Target_LetFron2_1580:=[[75.356,-99.732,84.333],[0.680036541,-0.521810391,-0.313535314,0.408607177],[0,0,0,0],[9E+09,9E+09,9E+09,9E+09,9E+09,9E+09]];
    CONST robtarget Target_LetFron2_1590:=[[76.129,-99.143,84.389],[0.680036541,-0.521810391,-0.313535314,0.408607177],[0,0,0,0],[9E+09,9E+09,9E+09,9E+09,9E+09,9E+09]];
    CONST robtarget Target_LetFron2_1600:=[[77.116,-98.378,84.254],[0.680036541,-0.521810391,-0.313535314,0.408607177],[0,0,0,0],[9E+09,9E+09,9E+09,9E+09,9E+09,9E+09]];
    CONST robtarget Target_LetFron2_1610:=[[78.006,-97.673,83.849],[0.680036541,-0.521810391,-0.313535314,0.408607177],[0,0,0,0],[9E+09,9E+09,9E+09,9E+09,9E+09,9E+09]];
    CONST robtarget Target_LetFron2_1620:=[[79.334,-96.597,82.185],[0.680036541,-0.521810391,-0.313535314,0.408607177],[0,0,0,0],[9E+09,9E+09,9E+09,9E+09,9E+09,9E+09]];
    CONST robtarget Target_LetFron2_1630:=[[79.82,-96.196,79.284],[0.680036541,-0.521810391,-0.313535314,0.408607177],[0,0,0,0],[9E+09,9E+09,9E+09,9E+09,9E+09,9E+09]];
    CONST robtarget Target_LetFron2_1640:=[[79.708,-96.29,77.625],[0.680036541,-0.521810391,-0.313535314,0.408607177],[0,0,0,0],[9E+09,9E+09,9E+09,9E+09,9E+09,9E+09]];
    CONST robtarget Target_LetFron2_1650:=[[79.369,-96.569,76.248],[0.680036541,-0.521810391,-0.313535314,0.408607177],[0,0,0,0],[9E+09,9E+09,9E+09,9E+09,9E+09,9E+09]];
    CONST robtarget Target_LetFron2_1660:=[[78.812,-97.024,75.146],[0.680036541,-0.521810391,-0.313535314,0.408607177],[0,0,0,0],[9E+09,9E+09,9E+09,9E+09,9E+09,9E+09]];
    CONST robtarget Target_LetFron2_1670:=[[78.077,-97.617,74.359],[0.680036541,-0.521810391,-0.313535314,0.408607177],[0,0,0,0],[9E+09,9E+09,9E+09,9E+09,9E+09,9E+09]];
    CONST robtarget Target_LetFron2_1680:=[[77.191,-98.319,73.87],[0.680036541,-0.521810391,-0.313535314,0.408607177],[0,0,0,0],[9E+09,9E+09,9E+09,9E+09,9E+09,9E+09]];
    CONST robtarget Target_LetFron2_1690:=[[75.499,-99.624,73.779],[0.680036541,-0.521810391,-0.313535314,0.408607177],[0,0,0,0],[9E+09,9E+09,9E+09,9E+09,9E+09,9E+09]];
    CONST robtarget Target_LetFron2_1700:=[[73.99,-100.75,74.808],[0.680036541,-0.521810391,-0.313535314,0.408607177],[0,0,0,0],[9E+09,9E+09,9E+09,9E+09,9E+09,9E+09]];
    CONST robtarget Target_LetFron2_1710:=[[73.426,-101.161,76.023],[0.680036541,-0.521810391,-0.313535314,0.408607177],[0,0,0,0],[9E+09,9E+09,9E+09,9E+09,9E+09,9E+09]];
    CONST robtarget Target_LetFron2_1720:=[[73.226,-101.306,77.552],[0.680036541,-0.521810391,-0.313535314,0.408607177],[0,0,0,0],[9E+09,9E+09,9E+09,9E+09,9E+09,9E+09]];
    CONST robtarget Target_LetFron2_1730:=[[73.281,-101.267,78.857],[0.680036541,-0.521810391,-0.313535314,0.408607177],[0,0,0,0],[9E+09,9E+09,9E+09,9E+09,9E+09,9E+09]];
    CONST robtarget Target_LetFron2_1740:=[[75.826,-99.375,78.857],[0.680036541,-0.521810391,-0.313535314,0.408607177],[0,0,0,0],[9E+09,9E+09,9E+09,9E+09,9E+09,9E+09]];
    CONST robtarget Target_LetFron2_1750:=[[78.322,-97.42,78.857],[0.680036541,-0.521810391,-0.313535314,0.408607177],[0,0,0,0],[9E+09,9E+09,9E+09,9E+09,9E+09,9E+09]];
    CONST robtarget Target_LetFron2_1760:=[[88.322,-117.42,78.857],[0.680036541,-0.521810391,-0.313535314,0.408607177],[0,0,0,0],[9E+09,9E+09,9E+09,9E+09,9E+09,9E+09]];
    CONST robtarget Target_LetFron2_1770:=[[90.513,-115.618,83.782],[0.680036541,-0.521810391,-0.313535314,0.408607177],[0,0,0,0],[9E+09,9E+09,9E+09,9E+09,9E+09,9E+09]];
    CONST robtarget Target_LetFron2_1780:=[[80.513,-95.618,83.782],[0.680036541,-0.521810391,-0.313535314,0.408607177],[0,0,0,0],[9E+09,9E+09,9E+09,9E+09,9E+09,9E+09]];
    CONST robtarget Target_LetFron2_1790:=[[83.101,-93.377,84.316],[0.680036541,-0.521810391,-0.313535314,0.408607177],[0,0,0,0],[9E+09,9E+09,9E+09,9E+09,9E+09,9E+09]];
    CONST robtarget Target_LetFron2_1800:=[[84.366,-92.235,83.242],[0.680036541,-0.521810391,-0.313535314,0.408607177],[0,0,0,0],[9E+09,9E+09,9E+09,9E+09,9E+09,9E+09]];
    CONST robtarget Target_LetFron2_1810:=[[84.565,-92.053,82.579],[0.680036541,-0.521810391,-0.313535314,0.408607177],[0,0,0,0],[9E+09,9E+09,9E+09,9E+09,9E+09,9E+09]];
    CONST robtarget Target_LetFron2_1820:=[[84.548,-92.068,72.267],[0.680036541,-0.521810391,-0.313535314,0.408607177],[0,0,0,0],[9E+09,9E+09,9E+09,9E+09,9E+09,9E+09]];
    CONST robtarget Target_LetFron2_1830:=[[84.565,-92.053,73.976],[0.680036541,-0.521810391,-0.313535314,0.408607177],[0,0,0,0],[9E+09,9E+09,9E+09,9E+09,9E+09,9E+09]];
    CONST robtarget Target_LetFron2_1840:=[[85.799,-90.904,74.201],[0.680036541,-0.521810391,-0.313535314,0.408607177],[0,0,0,0],[9E+09,9E+09,9E+09,9E+09,9E+09,9E+09]];
    CONST robtarget Target_LetFron2_1850:=[[80.667,-95.487,73.976],[0.680036541,-0.521810391,-0.313535314,0.408607177],[0,0,0,0],[9E+09,9E+09,9E+09,9E+09,9E+09,9E+09]];
    CONST robtarget Target_LetFron2_1860:=[[90.667,-115.487,73.976],[0.680036541,-0.521810391,-0.313535314,0.408607177],[0,0,0,0],[9E+09,9E+09,9E+09,9E+09,9E+09,9E+09]];
    CONST robtarget Target_LetFron2_1870:=[[97.066,-109.691,84.097],[0.680036541,-0.521810391,-0.313535314,0.408607177],[0,0,0,0],[9E+09,9E+09,9E+09,9E+09,9E+09,9E+09]];
    CONST robtarget Target_LetFron2_1880:=[[87.066,-89.691,84.097],[0.680036541,-0.521810391,-0.313535314,0.408607177],[0,0,0,0],[9E+09,9E+09,9E+09,9E+09,9E+09,9E+09]];
    CONST robtarget Target_LetFron2_1890:=[[87.066,-89.691,76.698],[0.680036541,-0.521810391,-0.313535314,0.408607177],[0,0,0,0],[9E+09,9E+09,9E+09,9E+09,9E+09,9E+09]];
    CONST robtarget Target_LetFron2_1900:=[[87.34,-89.425,75.101],[0.680036541,-0.521810391,-0.313535314,0.408607177],[0,0,0,0],[9E+09,9E+09,9E+09,9E+09,9E+09,9E+09]];
    CONST robtarget Target_LetFron2_1910:=[[87.669,-89.102,74.505],[0.680036541,-0.521810391,-0.313535314,0.408607177],[0,0,0,0],[9E+09,9E+09,9E+09,9E+09,9E+09,9E+09]];
    CONST robtarget Target_LetFron2_1920:=[[88.646,-88.13,73.796],[0.680036541,-0.521810391,-0.313535314,0.408607177],[0,0,0,0],[9E+09,9E+09,9E+09,9E+09,9E+09,9E+09]];
    CONST robtarget Target_LetFron2_1930:=[[89.643,-87.116,73.751],[0.680036541,-0.521810391,-0.313535314,0.408607177],[0,0,0,0],[9E+09,9E+09,9E+09,9E+09,9E+09,9E+09]];
    CONST robtarget Target_LetFron2_1940:=[[90.604,-86.116,74.156],[0.680036541,-0.521810391,-0.313535314,0.408607177],[0,0,0,0],[9E+09,9E+09,9E+09,9E+09,9E+09,9E+09]];
    CONST robtarget Target_LetFron2_1950:=[[91.579,-85.078,74.831],[0.680036541,-0.521810391,-0.313535314,0.408607177],[0,0,0,0],[9E+09,9E+09,9E+09,9E+09,9E+09,9E+09]];
    CONST robtarget Target_LetFron2_1960:=[[91.824,-84.814,73.706],[0.680036541,-0.521810391,-0.313535314,0.408607177],[0,0,0,0],[9E+09,9E+09,9E+09,9E+09,9E+09,9E+09]];
    CONST robtarget Target_LetFron2_1970:=[[92.295,-84.301,73.853],[0.680036541,-0.521810391,-0.313535314,0.408607177],[0,0,0,0],[9E+09,9E+09,9E+09,9E+09,9E+09,9E+09]];
    CONST robtarget Target_LetFron2_1980:=[[92.113,-84.5,84.097],[0.680036541,-0.521810391,-0.313535314,0.408607177],[0,0,0,0],[9E+09,9E+09,9E+09,9E+09,9E+09,9E+09]];
    CONST robtarget Target_LetFron2_1990:=[[102.113,-104.5,84.097],[0.680036541,-0.521810391,-0.313535314,0.408607177],[0,0,0,0],[9E+09,9E+09,9E+09,9E+09,9E+09,9E+09]];
    CONST robtarget Target_LetFron2_2000:=[[105.727,-100.382,84.097],[0.680036541,-0.521810391,-0.313535314,0.408607177],[0,0,0,0],[9E+09,9E+09,9E+09,9E+09,9E+09,9E+09]];
    CONST robtarget Target_LetFron2_2010:=[[95.727,-80.382,84.097],[0.680036541,-0.521810391,-0.313535314,0.408607177],[0,0,0,0],[9E+09,9E+09,9E+09,9E+09,9E+09,9E+09]];
    CONST robtarget Target_LetFron2_2020:=[[95.727,-80.382,70.333],[0.680036541,-0.521810391,-0.313535314,0.408607177],[0,0,0,0],[9E+09,9E+09,9E+09,9E+09,9E+09,9E+09]];
    CONST robtarget Target_LetFron2_2030:=[[105.727,-100.382,70.333],[0.680036541,-0.521810391,-0.313535314,0.408607177],[0,0,0,0],[9E+09,9E+09,9E+09,9E+09,9E+09,9E+09]];
    !***********************************************************
    !Dibujo el engranaje
    CONST robtarget Target_Frente_30:=[[-249.558695877,-44.184,-87.888947338],[0.695637986,0.547964836,-0.051631181,0.461688805],[0,-2,0,0],[9E+09,9E+09,9E+09,9E+09,9E+09,9E+09]];
    CONST robtarget Target_Frente_40:=[[-193.073509151,-40.184,-39.636157587],[0.522590279,0.416685464,0.130041044,0.732367361],[0,0,0,0],[9E+09,9E+09,9E+09,9E+09,9E+09,9E+09]];
    CONST robtarget Target_DibEng_10:=[[-147.685,-75.967,45.609],[0.589624104,0.343247558,0.546502531,0.485653697],[0,0,0,0],[9E+09,9E+09,9E+09,9E+09,9E+09,9E+09]];
    CONST robtarget Target_DibEng_20:=[[-137.628,-56.092,45.812],[0.589624104,0.343247558,0.546502531,0.485653697],[0,0,0,0],[9E+09,9E+09,9E+09,9E+09,9E+09,9E+09]];
    CONST robtarget Target_DibEng_30:=[[-137.654,-56.036,45.777],[0.589624104,0.343247558,0.546502531,0.485653697],[0,0,0,0],[9E+09,9E+09,9E+09,9E+09,9E+09,9E+09]];
    CONST robtarget Target_DibEng_40:=[[-138.241,-54.734,44.277],[0.589624104,0.343247558,0.546502531,0.485653697],[0,0,0,0],[9E+09,9E+09,9E+09,9E+09,9E+09,9E+09]];
    CONST robtarget Target_DibEng_50:=[[-138.766,-53.535,39.59],[0.589624104,0.343247558,0.546502531,0.485653697],[0,0,0,0],[9E+09,9E+09,9E+09,9E+09,9E+09,9E+09]];
    CONST robtarget Target_DibEng_60:=[[-140.069,-50.401,38.44],[0.589624104,0.343247558,0.546502531,0.485653697],[0,0,0,0],[9E+09,9E+09,9E+09,9E+09,9E+09,9E+09]];
    CONST robtarget Target_DibEng_70:=[[-141.468,-46.734,38.803],[0.589624104,0.343247558,0.546502531,0.485653697],[0,0,0,0],[9E+09,9E+09,9E+09,9E+09,9E+09,9E+09]];
    CONST robtarget Target_DibEng_80:=[[-141.886,-45.569,41.825],[0.589624104,0.343247558,0.546502531,0.485653697],[0,0,0,0],[9E+09,9E+09,9E+09,9E+09,9E+09,9E+09]];
    CONST robtarget Target_DibEng_90:=[[-142.007,-45.222,44.034],[0.589624104,0.343247558,0.546502531,0.485653697],[0,0,0,0],[9E+09,9E+09,9E+09,9E+09,9E+09,9E+09]];
    CONST robtarget Target_DibEng_100:=[[-142.434,-43.979,45.695],[0.589624104,0.343247558,0.546502531,0.485653697],[0,0,0,0],[9E+09,9E+09,9E+09,9E+09,9E+09,9E+09]];
    CONST robtarget Target_DibEng_110:=[[-143.128,-41.863,46.426],[0.589624104,0.343247558,0.546502531,0.485653697],[0,0,0,0],[9E+09,9E+09,9E+09,9E+09,9E+09,9E+09]];
    CONST robtarget Target_DibEng_120:=[[-143.616,-40.29,45.804],[0.589624104,0.343247558,0.546502531,0.485653697],[0,0,0,0],[9E+09,9E+09,9E+09,9E+09,9E+09,9E+09]];
    CONST robtarget Target_DibEng_130:=[[-144.199,-38.31,44.329],[0.589624104,0.343247558,0.546502531,0.485653697],[0,0,0,0],[9E+09,9E+09,9E+09,9E+09,9E+09,9E+09]];
    CONST robtarget Target_DibEng_140:=[[-144.768,-36.25,43.698],[0.589624104,0.343247558,0.546502531,0.485653697],[0,0,0,0],[9E+09,9E+09,9E+09,9E+09,9E+09,9E+09]];
    CONST robtarget Target_DibEng_150:=[[-145.419,-33.707,45.295],[0.589624104,0.343247558,0.546502531,0.485653697],[0,0,0,0],[9E+09,9E+09,9E+09,9E+09,9E+09,9E+09]];
    CONST robtarget Target_DibEng_160:=[[-145.898,-31.674,47.383],[0.589624104,0.343247558,0.546502531,0.485653697],[0,0,0,0],[9E+09,9E+09,9E+09,9E+09,9E+09,9E+09]];
    CONST robtarget Target_DibEng_170:=[[-145.932,-31.532,49.569],[0.589624104,0.343247558,0.546502531,0.485653697],[0,0,0,0],[9E+09,9E+09,9E+09,9E+09,9E+09,9E+09]];
    CONST robtarget Target_DibEng_180:=[[-145.711,-32.485,51.341],[0.589624104,0.343247558,0.546502531,0.485653697],[0,0,0,0],[9E+09,9E+09,9E+09,9E+09,9E+09,9E+09]];
    CONST robtarget Target_DibEng_190:=[[-145.368,-33.918,53.867],[0.589624104,0.343247558,0.546502531,0.485653697],[0,0,0,0],[9E+09,9E+09,9E+09,9E+09,9E+09,9E+09]];
    CONST robtarget Target_DibEng_200:=[[-145.42,-33.703,55.976],[0.589624104,0.343247558,0.546502531,0.485653697],[0,0,0,0],[9E+09,9E+09,9E+09,9E+09,9E+09,9E+09]];
    CONST robtarget Target_DibEng_210:=[[-145.914,-31.604,58.045],[0.589624104,0.343247558,0.546502531,0.485653697],[0,0,0,0],[9E+09,9E+09,9E+09,9E+09,9E+09,9E+09]];
    CONST robtarget Target_DibEng_220:=[[-146.605,-28.353,58.601],[0.589624104,0.343247558,0.546502531,0.485653697],[0,0,0,0],[9E+09,9E+09,9E+09,9E+09,9E+09,9E+09]];
    CONST robtarget Target_DibEng_230:=[[-146.95,-26.546,60.371],[0.589624104,0.343247558,0.546502531,0.485653697],[0,0,0,0],[9E+09,9E+09,9E+09,9E+09,9E+09,9E+09]];
    CONST robtarget Target_DibEng_240:=[[-146.992,-26.315,63.373],[0.589624104,0.343247558,0.546502531,0.485653697],[0,0,0,0],[9E+09,9E+09,9E+09,9E+09,9E+09,9E+09]];
    CONST robtarget Target_DibEng_250:=[[-146.9,-26.816,66.649],[0.589624104,0.343247558,0.546502531,0.485653697],[0,0,0,0],[9E+09,9E+09,9E+09,9E+09,9E+09,9E+09]];
    CONST robtarget Target_DibEng_260:=[[-146.507,-28.838,67.577],[0.589624104,0.343247558,0.546502531,0.485653697],[0,0,0,0],[9E+09,9E+09,9E+09,9E+09,9E+09,9E+09]];
    CONST robtarget Target_DibEng_270:=[[-145.997,-31.233,67.985],[0.589624104,0.343247558,0.546502531,0.485653697],[0,0,0,0],[9E+09,9E+09,9E+09,9E+09,9E+09,9E+09]];
    CONST robtarget Target_DibEng_280:=[[-145.58,-33.041,68.82],[0.589624104,0.343247558,0.546502531,0.485653697],[0,0,0,0],[9E+09,9E+09,9E+09,9E+09,9E+09,9E+09]];
    CONST robtarget Target_DibEng_290:=[[-145.402,-33.776,70.299],[0.589624104,0.343247558,0.546502531,0.485653697],[0,0,0,0],[9E+09,9E+09,9E+09,9E+09,9E+09,9E+09]];
    CONST robtarget Target_DibEng_300:=[[-145.395,-33.806,72.644],[0.589624104,0.343247558,0.546502531,0.485653697],[0,0,0,0],[9E+09,9E+09,9E+09,9E+09,9E+09,9E+09]];
    CONST robtarget Target_DibEng_310:=[[-145.874,-31.779,75.826],[0.589624104,0.343247558,0.546502531,0.485653697],[0,0,0,0],[9E+09,9E+09,9E+09,9E+09,9E+09,9E+09]];
    CONST robtarget Target_DibEng_320:=[[-145.991,-31.26,77.845],[0.589624104,0.343247558,0.546502531,0.485653697],[0,0,0,0],[9E+09,9E+09,9E+09,9E+09,9E+09,9E+09]];
    CONST robtarget Target_DibEng_330:=[[-145.641,-32.785,79.851],[0.589624104,0.343247558,0.546502531,0.485653697],[0,0,0,0],[9E+09,9E+09,9E+09,9E+09,9E+09,9E+09]];
    CONST robtarget Target_DibEng_340:=[[-145.309,-34.15,81.253],[0.589624104,0.343247558,0.546502531,0.485653697],[0,0,0,0],[9E+09,9E+09,9E+09,9E+09,9E+09,9E+09]];
    CONST robtarget Target_DibEng_350:=[[-144.767,-36.253,82.394],[0.589624104,0.343247558,0.546502531,0.485653697],[0,0,0,0],[9E+09,9E+09,9E+09,9E+09,9E+09,9E+09]];
    CONST robtarget Target_DibEng_360:=[[-144.225,-38.219,81.832],[0.589624104,0.343247558,0.546502531,0.485653697],[0,0,0,0],[9E+09,9E+09,9E+09,9E+09,9E+09,9E+09]];
    CONST robtarget Target_DibEng_370:=[[-143.564,-40.461,80.163],[0.589624104,0.343247558,0.546502531,0.485653697],[0,0,0,0],[9E+09,9E+09,9E+09,9E+09,9E+09,9E+09]];
    CONST robtarget Target_DibEng_380:=[[-142.961,-42.383,79.84],[0.589624104,0.343247558,0.546502531,0.485653697],[0,0,0,0],[9E+09,9E+09,9E+09,9E+09,9E+09,9E+09]];
    CONST robtarget Target_DibEng_390:=[[-142.434,-43.979,80.399],[0.589624104,0.343247558,0.546502531,0.485653697],[0,0,0,0],[9E+09,9E+09,9E+09,9E+09,9E+09,9E+09]];
    CONST robtarget Target_DibEng_400:=[[-142.133,-44.86,81.17],[0.589624104,0.343247558,0.546502531,0.485653697],[0,0,0,0],[9E+09,9E+09,9E+09,9E+09,9E+09,9E+09]];
    CONST robtarget Target_DibEng_410:=[[-141.772,-45.89,85.785],[0.589624104,0.343247558,0.546502531,0.485653697],[0,0,0,0],[9E+09,9E+09,9E+09,9E+09,9E+09,9E+09]];
    CONST robtarget Target_DibEng_420:=[[-141.531,-46.561,86.809],[0.589624104,0.343247558,0.546502531,0.485653697],[0,0,0,0],[9E+09,9E+09,9E+09,9E+09,9E+09,9E+09]];
    CONST robtarget Target_DibEng_430:=[[-141.029,-47.922,87.653],[0.589624104,0.343247558,0.546502531,0.485653697],[0,0,0,0],[9E+09,9E+09,9E+09,9E+09,9E+09,9E+09]];
    CONST robtarget Target_DibEng_440:=[[-139.311,-52.254,87.653],[0.589624104,0.343247558,0.546502531,0.485653697],[0,0,0,0],[9E+09,9E+09,9E+09,9E+09,9E+09,9E+09]];
    CONST robtarget Target_DibEng_450:=[[-138.658,-53.784,86.11],[0.589624104,0.343247558,0.546502531,0.485653697],[0,0,0,0],[9E+09,9E+09,9E+09,9E+09,9E+09,9E+09]];
    CONST robtarget Target_DibEng_460:=[[-138.45,-54.262,84.152],[0.589624104,0.343247558,0.546502531,0.485653697],[0,0,0,0],[9E+09,9E+09,9E+09,9E+09,9E+09,9E+09]];
    CONST robtarget Target_DibEng_470:=[[-138.242,-54.732,81.816],[0.589624104,0.343247558,0.546502531,0.485653697],[0,0,0,0],[9E+09,9E+09,9E+09,9E+09,9E+09,9E+09]];
    CONST robtarget Target_DibEng_480:=[[-137.623,-56.103,80.273],[0.589624104,0.343247558,0.546502531,0.485653697],[0,0,0,0],[9E+09,9E+09,9E+09,9E+09,9E+09,9E+09]];
    CONST robtarget Target_DibEng_490:=[[-136.745,-57.977,79.677],[0.589624104,0.343247558,0.546502531,0.485653697],[0,0,0,0],[9E+09,9E+09,9E+09,9E+09,9E+09,9E+09]];
    CONST robtarget Target_DibEng_500:=[[-136.285,-58.927,80.085],[0.589624104,0.343247558,0.546502531,0.485653697],[0,0,0,0],[9E+09,9E+09,9E+09,9E+09,9E+09,9E+09]];
    CONST robtarget Target_DibEng_510:=[[-135.75,-60.009,80.872],[0.589624104,0.343247558,0.546502531,0.485653697],[0,0,0,0],[9E+09,9E+09,9E+09,9E+09,9E+09,9E+09]];
    CONST robtarget Target_DibEng_520:=[[-135.067,-61.351,81.939],[0.589624104,0.343247558,0.546502531,0.485653697],[0,0,0,0],[9E+09,9E+09,9E+09,9E+09,9E+09,9E+09]];
    CONST robtarget Target_DibEng_530:=[[-134.488,-62.459,82.691],[0.589624104,0.343247558,0.546502531,0.485653697],[0,0,0,0],[9E+09,9E+09,9E+09,9E+09,9E+09,9E+09]];
    CONST robtarget Target_DibEng_540:=[[-133.661,-63.993,82.086],[0.589624104,0.343247558,0.546502531,0.485653697],[0,0,0,0],[9E+09,9E+09,9E+09,9E+09,9E+09,9E+09]];
    CONST robtarget Target_DibEng_550:=[[-132.142,-66.692,79.216],[0.589624104,0.343247558,0.546502531,0.485653697],[0,0,0,0],[9E+09,9E+09,9E+09,9E+09,9E+09,9E+09]];
    CONST robtarget Target_DibEng_560:=[[-131.802,-67.275,77.992],[0.589624104,0.343247558,0.546502531,0.485653697],[0,0,0,0],[9E+09,9E+09,9E+09,9E+09,9E+09,9E+09]];
    CONST robtarget Target_DibEng_570:=[[-131.8,-67.279,76.378],[0.589624104,0.343247558,0.546502531,0.485653697],[0,0,0,0],[9E+09,9E+09,9E+09,9E+09,9E+09,9E+09]];
    CONST robtarget Target_DibEng_580:=[[-132.186,-66.616,75.083],[0.589624104,0.343247558,0.546502531,0.485653697],[0,0,0,0],[9E+09,9E+09,9E+09,9E+09,9E+09,9E+09]];
    CONST robtarget Target_DibEng_590:=[[-132.639,-65.828,73.813],[0.589624104,0.343247558,0.546502531,0.485653697],[0,0,0,0],[9E+09,9E+09,9E+09,9E+09,9E+09,9E+09]];
    CONST robtarget Target_DibEng_600:=[[-133.002,-65.185,72.483],[0.589624104,0.343247558,0.546502531,0.485653697],[0,0,0,0],[9E+09,9E+09,9E+09,9E+09,9E+09,9E+09]];
    CONST robtarget Target_DibEng_610:=[[-132.985,-65.216,70.448],[0.589624104,0.343247558,0.546502531,0.485653697],[0,0,0,0],[9E+09,9E+09,9E+09,9E+09,9E+09,9E+09]];
    CONST robtarget Target_DibEng_620:=[[-132.429,-66.194,68.715],[0.589624104,0.343247558,0.546502531,0.485653697],[0,0,0,0],[9E+09,9E+09,9E+09,9E+09,9E+09,9E+09]];
    CONST robtarget Target_DibEng_630:=[[-132.047,-66.856,68.112],[0.589624104,0.343247558,0.546502531,0.485653697],[0,0,0,0],[9E+09,9E+09,9E+09,9E+09,9E+09,9E+09]];
    CONST robtarget Target_DibEng_640:=[[-129.82,-70.536,67.174],[0.589624104,0.343247558,0.546502531,0.485653697],[0,0,0,0],[9E+09,9E+09,9E+09,9E+09,9E+09,9E+09]];
    CONST robtarget Target_DibEng_650:=[[-129.022,-71.789,65.308],[0.589624104,0.343247558,0.546502531,0.485653697],[0,0,0,0],[9E+09,9E+09,9E+09,9E+09,9E+09,9E+09]];
    CONST robtarget Target_DibEng_660:=[[-129.022,-71.789,61.026],[0.589624104,0.343247558,0.546502531,0.485653697],[0,0,0,0],[9E+09,9E+09,9E+09,9E+09,9E+09,9E+09]];
    CONST robtarget Target_DibEng_670:=[[-129.311,-71.34,59.417],[0.589624104,0.343247558,0.546502531,0.485653697],[0,0,0,0],[9E+09,9E+09,9E+09,9E+09,9E+09,9E+09]];
    CONST robtarget Target_DibEng_680:=[[-130.015,-70.225,58.636],[0.589624104,0.343247558,0.546502531,0.485653697],[0,0,0,0],[9E+09,9E+09,9E+09,9E+09,9E+09,9E+09]];
    CONST robtarget Target_DibEng_690:=[[-132.072,-66.813,57.848],[0.589624104,0.343247558,0.546502531,0.485653697],[0,0,0,0],[9E+09,9E+09,9E+09,9E+09,9E+09,9E+09]];
    CONST robtarget Target_DibEng_700:=[[-132.926,-65.32,55.976],[0.589624104,0.343247558,0.546502531,0.485653697],[0,0,0,0],[9E+09,9E+09,9E+09,9E+09,9E+09,9E+09]];
    CONST robtarget Target_DibEng_710:=[[-133.117,-64.978,53.641],[0.589624104,0.343247558,0.546502531,0.485653697],[0,0,0,0],[9E+09,9E+09,9E+09,9E+09,9E+09,9E+09]];
    CONST robtarget Target_DibEng_720:=[[-131.923,-67.068,50.272],[0.589624104,0.343247558,0.546502531,0.485653697],[0,0,0,0],[9E+09,9E+09,9E+09,9E+09,9E+09,9E+09]];
    CONST robtarget Target_DibEng_730:=[[-131.795,-67.288,48.303],[0.589624104,0.343247558,0.546502531,0.485653697],[0,0,0,0],[9E+09,9E+09,9E+09,9E+09,9E+09,9E+09]];
    CONST robtarget Target_DibEng_740:=[[-132.581,-65.929,45.998],[0.589624104,0.343247558,0.546502531,0.485653697],[0,0,0,0],[9E+09,9E+09,9E+09,9E+09,9E+09,9E+09]];
    CONST robtarget Target_DibEng_750:=[[-134.078,-63.228,43.718],[0.589624104,0.343247558,0.546502531,0.485653697],[0,0,0,0],[9E+09,9E+09,9E+09,9E+09,9E+09,9E+09]];
    CONST robtarget Target_DibEng_760:=[[-134.96,-61.557,43.979],[0.589624104,0.343247558,0.546502531,0.485653697],[0,0,0,0],[9E+09,9E+09,9E+09,9E+09,9E+09,9E+09]];
    CONST robtarget Target_DibEng_770:=[[-136.663,-58.147,46.253],[0.589624104,0.343247558,0.546502531,0.485653697],[0,0,0,0],[9E+09,9E+09,9E+09,9E+09,9E+09,9E+09]];
    CONST robtarget Target_DibEng_780:=[[-137.598,-56.158,45.85],[0.589624104,0.343247558,0.546502531,0.485653697],[0,-1,0,0],[9E+09,9E+09,9E+09,9E+09,9E+09,9E+09]];
    CONST robtarget Target_DibEng_790:=[[-147.578,-76.202,45.875],[0.589624104,0.343247558,0.546502531,0.485653697],[0,-1,0,0],[9E+09,9E+09,9E+09,9E+09,9E+09,9E+09]];
    CONST robtarget Target_DibEng_800:=[[-150.412,-69.532,54.845],[0.664999268,0.432932025,0.478595617,0.375888375],[-1,0,-2,0],[9E+09,9E+09,9E+09,9E+09,9E+09,9E+09]];
    CONST robtarget Target_DibEng_810:=[[-140.384,-49.603,54.845],[0.664999268,0.432932025,0.478595617,0.375888375],[-1,0,-2,0],[9E+09,9E+09,9E+09,9E+09,9E+09,9E+09]];
    CONST robtarget Target_DibEng_820:=[[-141.369,-47.003,55.469],[0.664999268,0.432932025,0.478595617,0.375888375],[-1,0,-2,0],[9E+09,9E+09,9E+09,9E+09,9E+09,9E+09]];
    CONST robtarget Target_DibEng_830:=[[-142.259,-44.495,57.247],[0.664999268,0.432932025,0.478595617,0.375888375],[-1,0,-2,0],[9E+09,9E+09,9E+09,9E+09,9E+09,9E+09]];
    CONST robtarget Target_DibEng_840:=[[-142.794,-42.901,59.687],[0.664999268,0.432932025,0.478595617,0.375888375],[-1,0,-2,0],[9E+09,9E+09,9E+09,9E+09,9E+09,9E+09]];
    CONST robtarget Target_DibEng_850:=[[-143.005,-42.247,62.312],[0.664999268,0.432932025,0.478595617,0.375888375],[-1,0,-2,0],[9E+09,9E+09,9E+09,9E+09,9E+09,9E+09]];
    CONST robtarget Target_DibEng_860:=[[-142.87,-42.669,65.801],[0.664999268,0.432932025,0.478595617,0.375888375],[-1,0,-2,0],[9E+09,9E+09,9E+09,9E+09,9E+09,9E+09]];
    CONST robtarget Target_DibEng_870:=[[-142.469,-43.876,68.107],[0.664999268,0.432932025,0.478595617,0.375888375],[-1,0,-2,0],[9E+09,9E+09,9E+09,9E+09,9E+09,9E+09]];
    CONST robtarget Target_DibEng_880:=[[-141.592,-46.388,70.319],[0.664999268,0.432932025,0.478595617,0.375888375],[-1,0,-2,0],[9E+09,9E+09,9E+09,9E+09,9E+09,9E+09]];
    CONST robtarget Target_DibEng_890:=[[-140.518,-49.262,71.249],[0.664999268,0.432932025,0.478595617,0.375888375],[-1,0,-2,0],[9E+09,9E+09,9E+09,9E+09,9E+09,9E+09]];
    CONST robtarget Target_DibEng_900:=[[-138.895,-53.235,70.673],[0.664999268,0.432932025,0.478595617,0.375888375],[-1,0,-2,0],[9E+09,9E+09,9E+09,9E+09,9E+09,9E+09]];
    CONST robtarget Target_DibEng_910:=[[-138.076,-55.104,69.039],[0.664999268,0.432932025,0.478595617,0.375888375],[-1,0,-2,0],[9E+09,9E+09,9E+09,9E+09,9E+09,9E+09]];
    CONST robtarget Target_DibEng_920:=[[-137.114,-57.2,65.917],[0.664999268,0.432932025,0.478595617,0.375888375],[-1,0,-2,0],[9E+09,9E+09,9E+09,9E+09,9E+09,9E+09]];
    CONST robtarget Target_DibEng_930:=[[-136.991,-57.461,62.924],[0.664999268,0.432932025,0.478595617,0.375888375],[-1,0,-2,0],[9E+09,9E+09,9E+09,9E+09,9E+09,9E+09]];
    CONST robtarget Target_DibEng_940:=[[-137.114,-57.2,60.176],[0.664999268,0.432932025,0.478595617,0.375888375],[-1,0,-2,0],[9E+09,9E+09,9E+09,9E+09,9E+09,9E+09]];
    CONST robtarget Target_DibEng_950:=[[-138.096,-55.059,57.005],[0.664999268,0.432932025,0.478595617,0.375888375],[-1,0,-2,0],[9E+09,9E+09,9E+09,9E+09,9E+09,9E+09]];
    CONST robtarget Target_DibEng_960:=[[-138.922,-53.17,55.627],[0.664999268,0.432932025,0.478595617,0.375888375],[-1,0,-2,0],[9E+09,9E+09,9E+09,9E+09,9E+09,9E+09]];
    CONST robtarget Target_DibEng_970:=[[-139.596,-51.567,54.845],[0.664999268,0.432932025,0.478595617,0.375888375],[-1,0,-2,0],[9E+09,9E+09,9E+09,9E+09,9E+09,9E+09]];
    CONST robtarget Target_DibEng_980:=[[-140.412,-49.532,54.845],[0.664999268,0.432932025,0.478595617,0.375888375],[-1,0,-2,0],[9E+09,9E+09,9E+09,9E+09,9E+09,9E+09]];
    CONST robtarget Target_DibEng_990:=[[-150.405,-69.55,54.845],[0.664999268,0.432932025,0.478595617,0.375888375],[-1,0,-2,0],[9E+09,9E+09,9E+09,9E+09,9E+09,9E+09]];
    CONST robtarget Target_DibEng_1000:=[[-126.405,-65.55,-43.155],[0.600884572,0.356007489,0.53827741,0.471650112],[-1,0,-2,0],[9E+09,9E+09,9E+09,9E+09,9E+09,9E+09]];
    !***********************************************************
    !Dibujo tercer cuadrante de letrero frontal
    CONST robtarget Target_LetFron3_10:=[[-117.114,-108.644,45.956],[0.430645927,0.216920311,0.57802214,0.658316087],[0,0,0,0],[9E+09,9E+09,9E+09,9E+09,9E+09,9E+09]];
    CONST robtarget Target_LetFron3_20:=[[-107.122,-88.637,45.913],[0.430645927,0.216920311,0.57802214,0.658316087],[0,0,0,0],[9E+09,9E+09,9E+09,9E+09,9E+09,9E+09]];
    CONST robtarget Target_LetFron3_30:=[[-103.624,-91.909,45.113],[0.430645927,0.216920311,0.57802214,0.658316087],[0,0,0,0],[9E+09,9E+09,9E+09,9E+09,9E+09,9E+09]];
    CONST robtarget Target_LetFron3_40:=[[-103.083,-92.393,45.496],[0.430645927,0.216920311,0.57802214,0.658316087],[0,0,0,0],[9E+09,9E+09,9E+09,9E+09,9E+09,9E+09]];
    CONST robtarget Target_LetFron3_50:=[[-102.664,-92.764,46.069],[0.430645927,0.216920311,0.57802214,0.658316087],[0,0,0,0],[9E+09,9E+09,9E+09,9E+09,9E+09,9E+09]];
    CONST robtarget Target_LetFron3_60:=[[-102.441,-92.96,46.587],[0.430645927,0.216920311,0.57802214,0.658316087],[0,0,0,0],[9E+09,9E+09,9E+09,9E+09,9E+09,9E+09]];
    CONST robtarget Target_LetFron3_70:=[[-102.239,-93.137,47.586],[0.430645927,0.216920311,0.57802214,0.658316087],[0,0,0,0],[9E+09,9E+09,9E+09,9E+09,9E+09,9E+09]];
    CONST robtarget Target_LetFron3_80:=[[-102.227,-93.147,48.212],[0.430645927,0.216920311,0.57802214,0.658316087],[0,0,0,0],[9E+09,9E+09,9E+09,9E+09,9E+09,9E+09]];
    CONST robtarget Target_LetFron3_90:=[[-102.548,-92.866,49.153],[0.430645927,0.216920311,0.57802214,0.658316087],[0,0,0,0],[9E+09,9E+09,9E+09,9E+09,9E+09,9E+09]];
    CONST robtarget Target_LetFron3_100:=[[-102.965,-92.498,49.742],[0.430645927,0.216920311,0.57802214,0.658316087],[0,0,0,0],[9E+09,9E+09,9E+09,9E+09,9E+09,9E+09]];
    CONST robtarget Target_LetFron3_110:=[[-103.333,-92.17,50.056],[0.430645927,0.216920311,0.57802214,0.658316087],[0,0,0,0],[9E+09,9E+09,9E+09,9E+09,9E+09,9E+09]];
    CONST robtarget Target_LetFron3_120:=[[-104.061,-91.514,50.481],[0.430645927,0.216920311,0.57802214,0.658316087],[0,0,0,0],[9E+09,9E+09,9E+09,9E+09,9E+09,9E+09]];
    CONST robtarget Target_LetFron3_130:=[[-105.182,-90.482,51.085],[0.430645927,0.216920311,0.57802214,0.658316087],[0,0,0,0],[9E+09,9E+09,9E+09,9E+09,9E+09,9E+09]];
    CONST robtarget Target_LetFron3_140:=[[-105.719,-89.979,51.519],[0.430645927,0.216920311,0.57802214,0.658316087],[0,0,0,0],[9E+09,9E+09,9E+09,9E+09,9E+09,9E+09]];
    CONST robtarget Target_LetFron3_150:=[[-107.38,-88.386,52.197],[0.430645927,0.216920311,0.57802214,0.658316087],[0,0,0,0],[9E+09,9E+09,9E+09,9E+09,9E+09,9E+09]];
    CONST robtarget Target_LetFron3_160:=[[-107.289,-88.474,53.081],[0.430645927,0.216920311,0.57802214,0.658316087],[0,0,0,0],[9E+09,9E+09,9E+09,9E+09,9E+09,9E+09]];
    CONST robtarget Target_LetFron3_170:=[[-107.01,-88.746,53.872],[0.430645927,0.216920311,0.57802214,0.658316087],[0,0,0,0],[9E+09,9E+09,9E+09,9E+09,9E+09,9E+09]];
    CONST robtarget Target_LetFron3_180:=[[-106.537,-89.202,54.595],[0.430645927,0.216920311,0.57802214,0.658316087],[0,0,0,0],[9E+09,9E+09,9E+09,9E+09,9E+09,9E+09]];
    CONST robtarget Target_LetFron3_190:=[[-105.896,-89.812,55.029],[0.430645927,0.216920311,0.57802214,0.658316087],[0,0,0,0],[9E+09,9E+09,9E+09,9E+09,9E+09,9E+09]];
    CONST robtarget Target_LetFron3_200:=[[-105.02,-90.632,55.331],[0.430645927,0.216920311,0.57802214,0.658316087],[0,0,0,0],[9E+09,9E+09,9E+09,9E+09,9E+09,9E+09]];
    CONST robtarget Target_LetFron3_210:=[[-104.218,-91.37,55.384],[0.430645927,0.216920311,0.57802214,0.658316087],[0,0,0,0],[9E+09,9E+09,9E+09,9E+09,9E+09,9E+09]];
    CONST robtarget Target_LetFron3_220:=[[-103.326,-92.176,55.268],[0.430645927,0.216920311,0.57802214,0.658316087],[0,0,0,0],[9E+09,9E+09,9E+09,9E+09,9E+09,9E+09]];
    CONST robtarget Target_LetFron3_230:=[[-102.649,-92.777,55.055],[0.430645927,0.216920311,0.57802214,0.658316087],[0,0,0,0],[9E+09,9E+09,9E+09,9E+09,9E+09,9E+09]];
    CONST robtarget Target_LetFron3_240:=[[-102.042,-93.309,54.817],[0.430645927,0.216920311,0.57802214,0.658316087],[0,0,0,0],[9E+09,9E+09,9E+09,9E+09,9E+09,9E+09]];
    CONST robtarget Target_LetFron3_250:=[[-112.042,-113.309,54.814],[0.430645927,0.216920311,0.57802214,0.658316087],[0,0,0,0],[9E+09,9E+09,9E+09,9E+09,9E+09,9E+09]];
    CONST robtarget Target_LetFron3_260:=[[-108.858,-115.987,49.398],[0.430645927,0.216920311,0.57802214,0.658316087],[0,0,0,0],[9E+09,9E+09,9E+09,9E+09,9E+09,9E+09]];
    CONST robtarget Target_LetFron3_270:=[[-98.902,-95.951,49.397],[0.430645927,0.216920311,0.57802214,0.658316087],[0,0,0,0],[9E+09,9E+09,9E+09,9E+09,9E+09,9E+09]];
    CONST robtarget Target_LetFron3_280:=[[-97.309,-97.226,49.442],[0.430645927,0.216920311,0.57802214,0.658316087],[0,0,0,0],[9E+09,9E+09,9E+09,9E+09,9E+09,9E+09]];
    CONST robtarget Target_LetFron3_290:=[[-96.156,-98.122,49.772],[0.430645927,0.216920311,0.57802214,0.658316087],[0,0,0,0],[9E+09,9E+09,9E+09,9E+09,9E+09,9E+09]];
    CONST robtarget Target_LetFron3_300:=[[-95.374,-98.718,50.488],[0.430645927,0.216920311,0.57802214,0.658316087],[0,0,0,0],[9E+09,9E+09,9E+09,9E+09,9E+09,9E+09]];
    CONST robtarget Target_LetFron3_310:=[[-94.593,-99.304,51.741],[0.430645927,0.216920311,0.57802214,0.658316087],[0,0,0,0],[9E+09,9E+09,9E+09,9E+09,9E+09,9E+09]];
    CONST robtarget Target_LetFron3_320:=[[-94.39,-99.454,53.209],[0.430645927,0.216920311,0.57802214,0.658316087],[0,0,0,0],[9E+09,9E+09,9E+09,9E+09,9E+09,9E+09]];
    CONST robtarget Target_LetFron3_330:=[[-94.761,-99.179,54.352],[0.430645927,0.216920311,0.57802214,0.658316087],[0,0,0,0],[9E+09,9E+09,9E+09,9E+09,9E+09,9E+09]];
    CONST robtarget Target_LetFron3_340:=[[-95.636,-98.519,55.094],[0.430645927,0.216920311,0.57802214,0.658316087],[0,0,0,0],[9E+09,9E+09,9E+09,9E+09,9E+09,9E+09]];
    CONST robtarget Target_LetFron3_350:=[[-96.378,-97.951,55.401],[0.430645927,0.216920311,0.57802214,0.658316087],[0,0,0,0],[9E+09,9E+09,9E+09,9E+09,9E+09,9E+09]];
    CONST robtarget Target_LetFron3_360:=[[-97.78,-96.853,55.063],[0.430645927,0.216920311,0.57802214,0.658316087],[0,0,0,0],[9E+09,9E+09,9E+09,9E+09,9E+09,9E+09]];
    CONST robtarget Target_LetFron3_370:=[[-98.701,-96.114,54.468],[0.430645927,0.216920311,0.57802214,0.658316087],[0,0,0,0],[9E+09,9E+09,9E+09,9E+09,9E+09,9E+09]];
    CONST robtarget Target_LetFron3_380:=[[-98.924,-95.933,54.292],[0.430645927,0.216920311,0.57802214,0.658316087],[0,0,0,0],[9E+09,9E+09,9E+09,9E+09,9E+09,9E+09]];
    CONST robtarget Target_LetFron3_390:=[[-99.299,-95.627,55.259],[0.430645927,0.216920311,0.57802214,0.658316087],[0,0,0,0],[9E+09,9E+09,9E+09,9E+09,9E+09,9E+09]];
    CONST robtarget Target_LetFron3_400:=[[-100.358,-94.748,55.087],[0.430645927,0.216920311,0.57802214,0.658316087],[0,0,0,0],[9E+09,9E+09,9E+09,9E+09,9E+09,9E+09]];
    CONST robtarget Target_LetFron3_410:=[[-100.336,-94.766,47.788],[0.430645927,0.216920311,0.57802214,0.658316087],[0,0,0,0],[9E+09,9E+09,9E+09,9E+09,9E+09,9E+09]];
    CONST robtarget Target_LetFron3_420:=[[-100.094,-94.968,46.345],[0.430645927,0.216920311,0.57802214,0.658316087],[0,0,0,0],[9E+09,9E+09,9E+09,9E+09,9E+09,9E+09]];
    CONST robtarget Target_LetFron3_430:=[[-99.571,-95.402,45.441],[0.430645927,0.216920311,0.57802214,0.658316087],[0,0,0,0],[9E+09,9E+09,9E+09,9E+09,9E+09,9E+09]];
    CONST robtarget Target_LetFron3_440:=[[-98.556,-96.229,44.854],[0.430645927,0.216920311,0.57802214,0.658316087],[0,0,0,0],[9E+09,9E+09,9E+09,9E+09,9E+09,9E+09]];
    CONST robtarget Target_LetFron3_450:=[[-96.719,-97.687,44.801],[0.430645927,0.216920311,0.57802214,0.658316087],[0,0,0,0],[9E+09,9E+09,9E+09,9E+09,9E+09,9E+09]];
    CONST robtarget Target_LetFron3_460:=[[-95.557,-98.58,45.186],[0.430645927,0.216920311,0.57802214,0.658316087],[0,0,0,0],[9E+09,9E+09,9E+09,9E+09,9E+09,9E+09]];
    CONST robtarget Target_LetFron3_470:=[[-94.644,-99.266,45.6],[0.430645927,0.216920311,0.57802214,0.658316087],[0,0,0,0],[9E+09,9E+09,9E+09,9E+09,9E+09,9E+09]];
    CONST robtarget Target_LetFron3_480:=[[-94.949,-99.038,46.888],[0.430645927,0.216920311,0.57802214,0.658316087],[0,0,0,0],[9E+09,9E+09,9E+09,9E+09,9E+09,9E+09]];
    CONST robtarget Target_LetFron3_490:=[[-96.364,-97.962,46.428],[0.430645927,0.216920311,0.57802214,0.658316087],[0,0,0,0],[9E+09,9E+09,9E+09,9E+09,9E+09,9E+09]];
    CONST robtarget Target_LetFron3_500:=[[-97.392,-97.16,46.271],[0.430645927,0.216920311,0.57802214,0.658316087],[0,0,0,0],[9E+09,9E+09,9E+09,9E+09,9E+09,9E+09]];
    CONST robtarget Target_LetFron3_510:=[[-98.196,-96.521,46.443],[0.430645927,0.216920311,0.57802214,0.658316087],[0,0,0,0],[9E+09,9E+09,9E+09,9E+09,9E+09,9E+09]];
    CONST robtarget Target_LetFron3_520:=[[-98.708,-96.108,47.289],[0.430645927,0.216920311,0.57802214,0.658316087],[0,0,0,0],[9E+09,9E+09,9E+09,9E+09,9E+09,9E+09]];
    CONST robtarget Target_LetFron3_530:=[[-98.883,-95.966,48.272],[0.430645927,0.216920311,0.57802214,0.658316087],[0,0,0,0],[9E+09,9E+09,9E+09,9E+09,9E+09,9E+09]];
    CONST robtarget Target_LetFron3_540:=[[-98.902,-95.951,49.345],[0.430645927,0.216920311,0.57802214,0.658316087],[0,0,0,0],[9E+09,9E+09,9E+09,9E+09,9E+09,9E+09]];
    CONST robtarget Target_LetFron3_550:=[[-108.902,-115.951,49.38],[0.430645927,0.216920311,0.57802214,0.658316087],[0,0,0,0],[9E+09,9E+09,9E+09,9E+09,9E+09,9E+09]];
    CONST robtarget Target_LetFron3_560:=[[-102.646,-120.723,55.091],[0.430645927,0.216920311,0.57802214,0.658316087],[0,0,0,0],[9E+09,9E+09,9E+09,9E+09,9E+09,9E+09]];
    CONST robtarget Target_LetFron3_570:=[[-92.646,-100.723,55.09],[0.430645927,0.216920311,0.57802214,0.658316087],[0,0,0,0],[9E+09,9E+09,9E+09,9E+09,9E+09,9E+09]];
    CONST robtarget Target_LetFron3_580:=[[-92.61,-100.749,47.281],[0.430645927,0.216920311,0.57802214,0.658316087],[0,0,0,0],[9E+09,9E+09,9E+09,9E+09,9E+09,9E+09]];
    CONST robtarget Target_LetFron3_590:=[[-90.546,-102.19,44.719],[0.430645927,0.216920311,0.57802214,0.658316087],[0,0,0,0],[9E+09,9E+09,9E+09,9E+09,9E+09,9E+09]];
    CONST robtarget Target_LetFron3_600:=[[-87.122,-104.45,45.776],[0.430645927,0.216920311,0.57802214,0.658316087],[0,0,0,0],[9E+09,9E+09,9E+09,9E+09,9E+09,9E+09]];
